(* IEC 61131-3 sources: daoli-st-library/DL_Base (part 11) *)

(* ---- FB_DL_DutyStandbyRotation.st ---- *)
(*==============================================================================
 * 组件名称 (Component)  : FB_DL_DutyStandbyRotation
 * 所属子库 (Sublibrary) : DL_Base
 * 当前版本 (Version)    : 1.0.0
 * 兼容性   (Platform)   : CODESYS 3.5 / TwinCAT 3 / 汇川 InoProShop / Machine Expert
 *                         仅依赖 Standard.library（TON / R_TRIG / ABS），零厂商方言
 * 功能描述 (Function)   : 8 台泵 / 风机 / 压缩机的主备轮值与均衡调度。
 *                         按累计运行时间排序，把"需求台数"分给运行时间最短且满足启动条件
 *                         的机组；按周期把领机降为备机、备机升为领机；故障机立即跳过；
 *                         每台机受最小运行时长与最小停机时长双重保护，避免刚启就停把
 *                         接触器打烂；任何时刻不得把在运行的机组全部停掉。
 *                         解决多泵系统两类对立顽疾："永远只跑 1 号泵、2 号泵锈死"与
 *                         "轮值切得太勤、接触器与软启动器半年一换"。
 *
 * 【安全语义 / Safety semantics（编码侧不可弱化的四条）】
 *   1) 命令-反馈分离：本块只发启动命令（cmd 语义，FALSE = 停），运行状态一律以
 *      abUnitRunning 反馈为准，绝不假设"发了命令就等于在转"。
 *   2) 先启后停：停机放行条件是"目标集中已在运行的台数 >= 需求台数"，比"在运行台数
 *      >= 需求台数"更严。后者在换机场景下仍会短暂欠载（压力/流量掉一拍），本块刻意收紧。
 *   3) 故障机越权停机：abUnitFault = TRUE 且仍在运行时立即撤销命令，越过最小运行时长。
 *      这是最小运行时长保护的唯一例外。
 *   4) 无可用机组时（需求 > 0 且可用 = 0）已在运行的机组绝不因此被停——现场可能是
 *      就地/检修状态把"就绪"信号摘掉了，停掉正在供压的泵比少启一台危险得多。
 *
 * 【失真与语义披露 / Distortion disclosure】
 *   1) 运行时间账（afRunSec / auStartCount）是否断电保持由调用方决定（Retain 声明在
 *      调用侧）。不保持则每次上电从 0 起轮，轮值顺序每次开机都从 0 号机开始。
 *   2) 时间换算按 TIME 基准 1 ms（CODESYS / TwinCAT 3 / 汇川三平台一致）。移植到
 *      100 ns 基准平台时只需改 DL_DS_MS_PER_S 处的一行换算，逻辑不动。
 *   3) 按接口契约，参数冲突故障的复位沿会清零运行时间账——等同重置最小时长约束，
 *      复位前必须确认机组处于稳定工况（手册列为操作注意事项）。
 *   4) 排序为选择排序 O(64)。同运行时间的 tie-break 取"上一拍序列位置"而非索引升序：
 *      若死守索引升序，段 7 刚做完的轮值会在下一拍重新排序时被原样排回去，轮值等于
 *      永不生效（本批实测踩到的实现陷阱）。首扫序列为 0..7 恒等排列，因此冷启动行为
 *      与"索引升序"完全一致；轮值之后同值机组按轮值后的相对顺序排列，结果仍可复算。
 *
 * 开源溯源 (Origin)     : 原创实现（参考西门子 LBP 基础过程库中"最多 8 台聚合体"的粒度
 *                         与 cmd/ind 命令-反馈分离思想，以及 lead-lag 主备轮值工艺惯例，
 *                         clean-room 编写，未接触也未复制任何 LBP 源码）
 * 本文件内含       : TYPE  E_DL_RotationState（配套枚举，归属 DL_Base）
 *                    FB    FB_DL_DutyStandbyRotation
 * 依赖     (Depends)    : 无 DL_ 内部依赖；Standard.library: TON / R_TRIG
 * 红线自检 (Redline)    : R1 ✓ 零全局变量表与外部变量引用 ｜ R2 ✓ 零物理 IO 地址直写
 *                         R3 ✓ 纯 IEC 61131-3（定长数组 + 选择排序，无动态内存）
 *                         R4 ✓ 需求钳位 + 时间增量钳位 + 双向最小时长 + 计数饱和
 *                         R5 ✓ 全变量中英双语同行注释 ｜ R6 ✓ 四态 ENUM + CASE + ELSE 兜底
 *                         R7 ✓ 三实例主体最前部无条件刷新（本组件核心考点）
 * 修订历史 (Revision)   :
 *   2026-11-14  v1.0.0  首版入库（Phase 1 收口批次 · R3）
 *============================================================================*)

(*-----------------------------------------------------------------------------
 * 枚举: E_DL_RotationState（归属 DL_Base，与 FB_DL_DutyStandbyRotation 同文件）
 * 含义: 轮值调度主状态。数值步长留空位便于后续插态而不破坏已有工程。
 *----------------------------------------------------------------------------*)
TYPE E_DL_RotationState :
(
    eIdle          := 0,     // 未使能：命令全部撤销，运行时间账继续按反馈累加 / Disabled, commands dropped, runtime still accounted
    eRunning       := 10,    // 正常调度：累加 → 排序 → 定需求集 → 先启后停 / Normal scheduling
    eRotatePending := 20,    // 轮值挂起：受最小时长阻挡，保持当前组合并每拍重试 / Rotation pending, retried every scan
    eFault         := 99     // 参数冲突锁存：轮值禁用，但启停调度照常工作 / Latched config fault, scheduling still runs
);
END_TYPE

(*==============================================================================
 * 功能块: FB_DL_DutyStandbyRotation
 * 调用约定: 每个扫描周期无条件调用一次，uDeltaTimeMs 必须注入真实任务间隔。
 *============================================================================*)
FUNCTION_BLOCK FB_DL_DutyStandbyRotation
VAR_INPUT
    abUnitReady     : ARRAY[0..7] OF BOOL;    // 机组就绪（无故障、无就地、无禁止），上限 8 台 / Unit ready, max 8 units
    abUnitRunning   : ARRAY[0..7] OF BOOL;    // 运行反馈（接触器辅助触点或流量开关）/ Running feedback
    abUnitFault     : ARRAY[0..7] OF BOOL;    // 机组故障（跳过并允许立即停机）/ Unit fault, skipped and stopped at once
    nDemand         : INT := 0;               // 需求运行台数，合法域 0..8 / Required unit count, valid 0..8
    bEnable         : BOOL := TRUE;           // 使能，FALSE 时命令全撤 / Enable, FALSE drops all commands
    uDeltaTimeMs    : UDINT;                  // 调用方注入的扫描间隔 [ms] / Injected scan delta [ms]
    tMinRunTime     : TIME := T#10M;          // 最小连续运行时长 [min]，防刚启就停 / Minimum run time
    tMinStopTime    : TIME := T#5M;           // 最小停机时长 [min]，防接触器高频动作 / Minimum stop time
    tRotateInterval : TIME := T#24H;          // 轮值周期 [h] / Rotation interval
    bForceRotate    : BOOL;                   // 上升沿：立即请求一次轮值（仍受最小时长约束）/ Rising edge: force one rotation
    bReset          : BOOL;                   // 上升沿：复位参数冲突并清零运行时间账 / Rising edge: reset the config fault and clear runtimes
END_VAR
VAR_OUTPUT
    abStartCmd        : ARRAY[0..7] OF BOOL;  // 启动命令（cmd 语义，FALSE = 停）/ Start command per unit, FALSE = stop
    anRank            : ARRAY[0..7] OF INT;   // 本轮优先顺序，0 = 最高 / Priority rank, 0 = highest
    nLeadUnit         : INT;                  // 领机号 0..7，-1 = 无 / Lead unit 0..7, -1 = none
    afRuntimeHours    : ARRAY[0..7] OF LREAL; // 累计运行小时 [h] / Accumulated runtime [h]
    abBlockedByMinRun : ARRAY[0..7] OF BOOL;  // 因最小运行时长被阻止停机 / Stop blocked by the minimum run time
    abBlockedByMinStop: ARRAY[0..7] OF BOOL;  // 因最小停机时长被阻止启动 / Start blocked by the minimum stop time
    auStartCount      : ARRAY[0..7] OF UDINT; // 各机启动次数（饱和）/ Start count per unit, saturating
    bRotatePending    : BOOL;                 // 轮值挂起中 / Rotation pending
    bNoAvailableUnit  : BOOL;                 // 无可用机组（瞬时诊断）/ No available unit, instantaneous
    uRotateCount      : UDINT;                // 已完成的轮值次数（饱和）/ Completed rotations, saturating
    bError            : BOOL;                 // 故障标志（参数冲突锁存）/ Fault flag, config conflict latched
    uErrorId          : UDINT;                // 故障码，0 = 无故障 / Error code, 0 = no error
    eState            : E_DL_RotationState;   // 当前状态（供 HMI 诊断）/ Current state for HMI diagnosis
END_VAR
VAR
    fbTrigReset     : R_TRIG;                 // 复位上升沿检测实例 / Reset rising edge detector
    fbTrigForce     : R_TRIG;                 // 强制轮值上升沿检测实例 / Force-rotate rising edge detector
    fbTonRotate     : TON;                    // 轮值周期定时器 / Rotation interval timer
    eStateInt       : E_DL_RotationState;     // 主状态机内部当前态 / Internal state of the main state machine
    afRunSec        : ARRAY[0..7] OF LREAL;   // 运行秒累加 [s] / Runtime seconds accumulator [s]
    afStopSec       : ARRAY[0..7] OF LREAL;   // 停机秒累加 [s] / Stop seconds accumulator [s]
    anOrder         : ARRAY[0..7] OF INT;     // 已提交的优先序列（可用优先，运行时间升序）/ Committed priority order
    anTrial         : ARRAY[0..7] OF INT;     // 轮值试验序列（未提交前不生效）/ Trial order, not committed yet
    anPos           : ARRAY[0..7] OF INT;     // 各机组在上一拍序列中的位置（排序稳定性锚点）/ Previous position per unit
    abUsable        : ARRAY[0..7] OF BOOL;    // 可用 = 就绪且无故障 / Usable = ready and not faulted
    abDesired       : ARRAY[0..7] OF BOOL;    // 目标运行集 / Desired running set
    abTrialUnit     : ARRAY[0..7] OF BOOL;    // 轮值试验目标集 / Trial desired set
    abCmdInt        : ARRAY[0..7] OF BOOL;    // 本拍命令内部副本 / Internal command copy of this scan
    abCmdPrev       : ARRAY[0..7] OF BOOL;    // 上一拍命令（算启动沿）/ Previous commands, for start edges
    nIdx            : INT;                    // 外层索引 / Outer index
    nInner          : INT;                    // 内层索引 / Inner index
    nMinPos         : INT;                    // 选择排序中的最小元位置 / Position of the minimum during selection sort
    nTmp            : INT;                    // 交换临时量 / Swap temporary
    nAvail          : INT;                    // 可用机组数 / Number of usable units
    nDesired        : INT;                    // 本拍应运行台数（已按可用数钳位）/ Desired count, clamped to the usable count
    nRunningCnt     : INT;                    // 当前在运行台数 / Currently running units
    nDesiredRunning : INT;                    // 目标集中已在运行的台数 / Desired units already running
    nCnt            : INT;                    // 计数累加器 / Counting accumulator
    nLead           : INT;                    // 领机号 / Lead unit index
    nDemandEff      : INT;                    // 钳位后的需求台数 / Clamped demand
    fDtSec          : LREAL;                  // 扫描间隔换算成秒 [s] / Scan delta in seconds [s]
    fMinRunSec      : LREAL;                  // 最小运行时长 [s] / Minimum run time [s]
    fMinStopSec     : LREAL;                  // 最小停机时长 [s] / Minimum stop time [s]
    tRotEff         : TIME;                   // 钳位后的轮值周期 [ms] / Clamped rotation interval [ms]
    uDtEff          : UDINT;                  // 钳位后的扫描间隔 [ms] / Clamped scan delta [ms]
    uWarnId         : UDINT;                  // 本拍瞬时告警码 / Instantaneous warning code of this scan
    uRotateCnt      : UDINT;                  // 轮值次数内部副本（饱和）/ Internal rotation counter, saturating
    bRotateReq      : BOOL;                   // 本拍请求轮值 / Rotation requested this scan
    bRotTimerRun    : BOOL;                   // 轮值定时器运行中 / Rotation timer running
    bRotTimerRearm  : BOOL;                   // 轮值定时器下一拍重新计时 / Rearm the rotation timer next scan
    bRotPendingScr  : BOOL;                   // 本拍轮值因最小时长受阻 / Rotation blocked by the minimum times this scan
    bFeasible       : BOOL;                   // 轮值试验是否可行 / Whether the trial rotation is feasible
    bSmaller        : BOOL;                   // 排序比较：候选元是否更靠前 / Sort comparator: candidate ranks earlier
    bHoldAll        : BOOL;                   // 无可用机组时冻结全部停机 / Freeze every stop when no unit is usable
    bSchedOn        : BOOL;                   // 本拍允许调度 / Scheduling enabled this scan
    bConflict       : BOOL;                   // 本拍存在时间参数冲突 / Time-parameter conflict present this scan
    bParamLatch     : BOOL;                   // 参数冲突锁存 / Configuration conflict latched
    bStateFault     : BOOL;                   // 非法状态锁存（与参数冲突分开记账）/ Illegal-state latch, kept apart from the config latch
    bCntWarned      : BOOL;                   // 饱和告警已发过一次 / Saturation warning already raised
    bSortInit       : BOOL := TRUE;           // 排序序列尚未初始化为恒等排列 / Priority order not yet initialised
    bFirstScan      : BOOL := TRUE;           // 上电首扫标志 / First-scan flag
END_VAR
VAR CONSTANT
    DL_DS_UNITS      : INT   := 8;            // 机组数，必须等于数组维度 / Unit count, must match the arrays
    DL_DS_IDX_NONE   : INT   := -1;           // 无效索引哨兵 / Invalid-index sentinel
    DL_DS_HOUR_MAX   : LREAL := 1.0E9;        // 运行小时饱和上限 [h] / Runtime saturation [h]
    DL_DS_SEC_MAX    : LREAL := 3.6E12;       // 运行秒饱和上限 [s]，与小时上限对齐 / Runtime saturation [s]
    DL_DS_SEC_PER_H  : LREAL := 3600.0;       // 小时换算常数 [s/h] / Seconds per hour
    DL_DS_MS_PER_S   : LREAL := 1000.0;       // 毫秒换算常数 [ms/s]，三平台 TIME 基准均为 1 ms / Milliseconds per second
    DL_DS_DT_MAX     : UDINT := 60000;        // 时间增量上限 [ms]，超此值判为断点 / Delta clamp [ms]
    DL_DS_EPS        : LREAL := 1.0E-6;       // 浮点判等容差 / Float comparison tolerance
    DL_DS_CNT_MAX    : UDINT := 16#FFFF_FFFE; // 计数器饱和值 / Counter saturation
    DL_DS_ROT_MIN    : TIME  := T#1S;         // 轮值周期下限 [s] / Rotation interval lower bound
    DL_DS_ROT_MAX    : TIME  := T#8760H;      // 轮值周期上限 [h]，一年 / Rotation interval upper bound
END_VAR

(*------------------------------------------------------------------------------
 * 段 0｜轮值周期钳位（先于定时器，避免 PT = 0 造成每拍触发）
 *      Rotation-interval clamp, done before the timer so PT is never zero
 *-----------------------------------------------------------------------------*)
uWarnId := 16#0000;
tRotEff := tRotateInterval;

IF tRotEff < DL_DS_ROT_MIN THEN
    tRotEff := DL_DS_ROT_MIN;
    uWarnId := 16#0001_0001;
ELSIF tRotEff > DL_DS_ROT_MAX THEN
    tRotEff := DL_DS_ROT_MAX;
    uWarnId := 16#0001_0001;
END_IF

(*------------------------------------------------------------------------------
 * 段 1｜无条件刷新区（红线 R7）：两沿 + 一轮值周期计时
 *      Unconditional refresh zone: two edges plus the rotation interval timer
 *      IN 由 bRotTimerRun 这一派生量给出，实例调用本身绝不进 IF
 *-----------------------------------------------------------------------------*)
fbTrigReset(CLK := bReset);
fbTrigForce(CLK := bForceRotate);
fbTonRotate(IN := bRotTimerRun, PT := tRotEff);

bRotateReq := fbTrigForce.Q;

IF fbTonRotate.Q THEN
    bRotateReq     := TRUE;
    bRotTimerRun   := FALSE;    // 下一拍 ET 归零 / Reset ET on the next scan
    bRotTimerRearm := TRUE;
ELSIF bRotTimerRearm THEN
    bRotTimerRun   := TRUE;
    bRotTimerRearm := FALSE;
END_IF

(*------------------------------------------------------------------------------
 * 段 2｜上电首扫：状态、领机号与锁存显式落到安全侧
 *      First-scan init: state, lead index and latches forced to the safe side
 *-----------------------------------------------------------------------------*)
IF bFirstScan THEN
    bFirstScan  := FALSE;
    eStateInt   := E_DL_RotationState.eIdle;
    nLead       := DL_DS_IDX_NONE;
    bParamLatch := FALSE;
    uRotateCnt  := 0;
    bRotTimerRun   := FALSE;
    bRotTimerRearm := TRUE;
END_IF

(*------------------------------------------------------------------------------
 * 段 3｜时间增量校验（边界 B8）：0 或超上限一律钳位，绝不接受回绕值
 *      Delta-time check: zero or over-limit values are clamped, wraparound never accepted
 *      回绕的 UDINT 转成秒后是天文数字，会瞬间把运行时间算爆并把排序彻底打乱
 *-----------------------------------------------------------------------------*)
IF uDeltaTimeMs = 0 THEN
    uDtEff  := 1;
    uWarnId := 16#0001_0008;
ELSIF uDeltaTimeMs > DL_DS_DT_MAX THEN
    uDtEff  := DL_DS_DT_MAX;
    uWarnId := 16#0001_0008;
ELSE
    uDtEff := uDeltaTimeMs;
END_IF

fDtSec     := UDINT_TO_LREAL(uDtEff) / DL_DS_MS_PER_S;
fMinRunSec := TIME_TO_LREAL(tMinRunTime) / DL_DS_MS_PER_S;
fMinStopSec := TIME_TO_LREAL(tMinStopTime) / DL_DS_MS_PER_S;

(*------------------------------------------------------------------------------
 * 段 4｜参数校验（边界 B1/B7）
 *      Parameter validation: demand clamp and the minimum-time conflict check
 *-----------------------------------------------------------------------------*)
nDemandEff := nDemand;
IF nDemand < 0 THEN
    nDemandEff := 0;
    uWarnId    := 16#0001_0001;
ELSIF nDemand > DL_DS_UNITS THEN
    nDemandEff := DL_DS_UNITS;
    uWarnId    := 16#0001_0001;
END_IF

(* 最小运行 + 最小停机 > 轮值周期：轮值永远等不到，属参数冲突而非运行故障 *)
(* min-run + min-stop > interval means rotation could never complete: a configuration conflict *)
bConflict := ((tMinRunTime + tMinStopTime) > tRotateInterval);

IF bConflict THEN
    bParamLatch := TRUE;
END_IF

IF (tMinRunTime < T#0S) OR (tMinStopTime < T#0S) THEN
    uWarnId := 16#0001_0001;
END_IF

(*------------------------------------------------------------------------------
 * 段 5｜运行时间记账（状态 eIdle 也照记：停机也要记账，否则轮值失真）
 *      Runtime accounting runs even when disabled: an unaccounted stop skews rotation
 *      以反馈为准而不是以命令为准，接触器没吸合就不能算运行
 *-----------------------------------------------------------------------------*)
FOR nIdx := 0 TO (DL_DS_UNITS - 1) DO

    IF abUnitRunning[nIdx] THEN
        afRunSec[nIdx] := afRunSec[nIdx] + fDtSec;
        IF afRunSec[nIdx] > DL_DS_SEC_MAX THEN
            afRunSec[nIdx] := DL_DS_SEC_MAX;
            uWarnId := 16#0001_0007;
        END_IF
    ELSE
        afStopSec[nIdx] := afStopSec[nIdx] + fDtSec;
        IF afStopSec[nIdx] > DL_DS_SEC_MAX THEN
            afStopSec[nIdx] := DL_DS_SEC_MAX;
        END_IF
    END_IF

    afRuntimeHours[nIdx] := afRunSec[nIdx] / DL_DS_SEC_PER_H;
    IF afRuntimeHours[nIdx] > DL_DS_HOUR_MAX THEN
        afRuntimeHours[nIdx] := DL_DS_HOUR_MAX;
    END_IF

END_FOR

(*------------------------------------------------------------------------------
 * 段 6｜可用性与候选排序（边界 B6/B10）
 *      Usability and candidate ordering: usable first, then runtime, then previous position
 *      序列只在首扫初始化为恒等排列，之后一律在既有排列上就地排序：
 *      若每拍都从 0..7 重新开始排，段 7 刚做完的轮值会在下一拍被排序抹掉，
 *      轮值等于永远不生效——这是本组件最容易踩的实现陷阱
 *      The order is initialised once and then sorted in place, otherwise every rotation
 *      would be erased by the next scan's re-sort
 *-----------------------------------------------------------------------------*)
nAvail := 0;

FOR nIdx := 0 TO (DL_DS_UNITS - 1) DO
    abUsable[nIdx] := abUnitReady[nIdx] AND (NOT abUnitFault[nIdx]);
    IF abUsable[nIdx] THEN
        nAvail := nAvail + 1;
    END_IF
END_FOR

IF bSortInit THEN
    FOR nIdx := 0 TO (DL_DS_UNITS - 1) DO
        anOrder[nIdx] := nIdx;
        anPos[nIdx]   := nIdx;
    END_FOR
    bSortInit := FALSE;
END_IF

(* 选择排序：8 元定长，0..6 外层、nIdx+1..7 内层，迭代次数由常量卡死 *)
(* Selection sort over 8 fixed elements, the loop bounds are compile-time constants *)
FOR nIdx := 0 TO (DL_DS_UNITS - 2) DO

    nMinPos := nIdx;

    FOR nInner := (nIdx + 1) TO (DL_DS_UNITS - 1) DO

        bSmaller := FALSE;

        IF abUsable[anOrder[nInner]] AND (NOT abUsable[anOrder[nMinPos]]) THEN
            bSmaller := TRUE;
        ELSIF abUsable[anOrder[nInner]] = abUsable[anOrder[nMinPos]] THEN
            IF (afRunSec[anOrder[nInner]] + DL_DS_EPS) < afRunSec[anOrder[nMinPos]] THEN
                bSmaller := TRUE;
            ELSIF ABS(afRunSec[anOrder[nInner]] - afRunSec[anOrder[nMinPos]]) <= DL_DS_EPS THEN
                (* 运行时间相同：按上一拍位置排序，保证稳定且轮值结果不被抹掉 *)
                (* Equal runtime: keep the previous relative order, so rotations survive *)
                IF anPos[anOrder[nInner]] < anPos[anOrder[nMinPos]] THEN
                    bSmaller := TRUE;
                END_IF
            END_IF
        END_IF

        IF bSmaller THEN
            nMinPos := nInner;
        END_IF

    END_FOR

    IF nMinPos <> nIdx THEN
        nTmp             := anOrder[nIdx];
        anOrder[nIdx]    := anOrder[nMinPos];
        anOrder[nMinPos] := nTmp;
    END_IF

END_FOR

FOR nIdx := 0 TO (DL_DS_UNITS - 1) DO
    anPos[anOrder[nIdx]] := nIdx;
END_FOR

nDesired := nDemandEff;
IF nDesired > nAvail THEN
    nDesired := nAvail;
END_IF

(*------------------------------------------------------------------------------
 * 段 7｜轮值尝试（边界 B7）：可行才移位，不可行一律不动任何命令
 *      Rotation attempt: shift only when every constraint is met, never touch commands otherwise
 *      把"领机移到可用序列末位、其余前移一位"这一动作做成试验序列，
 *      可行性由"要停的机组已满足最小运行、要启的机组已满足最小停机"共同决定
 *-----------------------------------------------------------------------------*)
bRotPendingScr := FALSE;

FOR nIdx := 0 TO (DL_DS_UNITS - 1) DO
    abBlockedByMinRun[nIdx]  := FALSE;
    abBlockedByMinStop[nIdx] := FALSE;
END_FOR

IF bRotateReq AND bEnable AND (NOT bParamLatch)
   AND (eStateInt <> E_DL_RotationState.eIdle)
   AND (eStateInt <> E_DL_RotationState.eFault)
   AND (nAvail >= 2) AND (nDesired >= 1) THEN

    FOR nIdx := 0 TO (DL_DS_UNITS - 1) DO
        anTrial[nIdx] := anOrder[nIdx];
    END_FOR

    nTmp := anTrial[0];
    FOR nIdx := 0 TO (DL_DS_UNITS - 2) DO
        IF nIdx < (nAvail - 1) THEN
            anTrial[nIdx] := anTrial[nIdx + 1];
        END_IF
    END_FOR
    anTrial[nAvail - 1] := nTmp;

    (* 试验目标集：可用序列中取前 nDesired 台 *)
    (* Trial set: the first nDesired usable entries of the trial order *)
    FOR nIdx := 0 TO (DL_DS_UNITS - 1) DO
        abTrialUnit[nIdx] := FALSE;
    END_FOR

    nCnt := 0;
    FOR nIdx := 0 TO (DL_DS_UNITS - 1) DO
        IF (nCnt < nDesired) AND abUsable[anTrial[nIdx]] AND (NOT abTrialUnit[anTrial[nIdx]]) THEN
            abTrialUnit[anTrial[nIdx]] := TRUE;
            nCnt := nCnt + 1;
        END_IF
    END_FOR

    (* 可行性检查：需停的看最小运行，需启的看最小停机；故障机不参与（越权立即停） *)
    (* Feasibility: stops need the min run time, starts need the min stop time *)
    bFeasible := TRUE;

    FOR nIdx := 0 TO (DL_DS_UNITS - 1) DO
        IF abUnitRunning[nIdx] AND (NOT abTrialUnit[nIdx]) AND (NOT abUnitFault[nIdx]) THEN
            IF afRunSec[nIdx] < fMinRunSec THEN
                bFeasible := FALSE;
                abBlockedByMinRun[nIdx] := TRUE;
            END_IF
        END_IF
        IF (NOT abUnitRunning[nIdx]) AND abTrialUnit[nIdx] THEN
            IF afStopSec[nIdx] < fMinStopSec THEN
                bFeasible := FALSE;
                abBlockedByMinStop[nIdx] := TRUE;
            END_IF
        END_IF
    END_FOR

    IF bFeasible THEN
        FOR nIdx := 0 TO (DL_DS_UNITS - 1) DO
            anOrder[nIdx] := anTrial[nIdx];
        END_FOR
        (* 提交后立即刷新位置锚点，否则下一次排序会按旧位置把轮值结果排回去 *)
        (* Refresh the position anchor at once, or the next sort undoes the rotation *)
        FOR nIdx := 0 TO (DL_DS_UNITS - 1) DO
            anPos[anOrder[nIdx]] := nIdx;
        END_FOR
        bRotateReq := FALSE;
        IF uRotateCnt < DL_DS_CNT_MAX THEN
            uRotateCnt := uRotateCnt + 1;
        ELSIF NOT bCntWarned THEN
            uWarnId    := 16#0001_0007;
            bCntWarned := TRUE;
        END_IF
    ELSE
        (* 边界 B7：请求不丢，保留到条件满足，每拍重试且只补做一次 *)
        (* The request is kept, retried every scan, and only ever executed once *)
        bRotPendingScr := TRUE;
    END_IF

END_IF

(*------------------------------------------------------------------------------
 * 段 8｜主状态机（红线 R6）：ENUM + CASE + ELSE 兜底
 *      Main state machine with the mandatory ELSE fallback
 *-----------------------------------------------------------------------------*)
CASE eStateInt OF

    E_DL_RotationState.eIdle:
        bRotateReq     := FALSE;
        bRotTimerRun   := FALSE;
        bRotTimerRearm := TRUE;
        IF bEnable THEN
            IF bParamLatch THEN
                eStateInt := E_DL_RotationState.eFault;
            ELSE
                eStateInt := E_DL_RotationState.eRunning;
            END_IF
        END_IF

    E_DL_RotationState.eRunning:
        IF NOT bEnable THEN
            eStateInt := E_DL_RotationState.eIdle;
        ELSIF bParamLatch THEN
            eStateInt := E_DL_RotationState.eFault;
        ELSIF bRotPendingScr THEN
            eStateInt := E_DL_RotationState.eRotatePending;
        END_IF

    E_DL_RotationState.eRotatePending:
        IF NOT bEnable THEN
            eStateInt := E_DL_RotationState.eIdle;
        ELSIF bParamLatch THEN
            eStateInt := E_DL_RotationState.eFault;
        ELSIF NOT bRotPendingScr THEN
            eStateInt := E_DL_RotationState.eRunning;
        END_IF

    E_DL_RotationState.eFault:
        (* 轮值禁用但启停调度照常：不能因为轮值配错就让泵不转 *)
        (* Rotation is disabled, scheduling still runs: a wrong interval must not stop the pumps *)
        bRotateReq := FALSE;
        IF NOT bEnable THEN
            eStateInt := E_DL_RotationState.eIdle;
        ELSIF fbTrigReset.Q AND (NOT bConflict) THEN
            bParamLatch := FALSE;
            bStateFault := FALSE;
            eStateInt   := E_DL_RotationState.eRunning;
            (* 接口契约：复位参数冲突同时清零运行时间账，等同重置最小时长约束 *)
            (* Contract: resetting the conflict also clears the runtime books *)
            FOR nIdx := 0 TO (DL_DS_UNITS - 1) DO
                afRunSec[nIdx]    := 0.0;
                afStopSec[nIdx]   := 0.0;
                afRuntimeHours[nIdx] := 0.0;
            END_FOR
            bRotTimerRun   := FALSE;
            bRotTimerRearm := TRUE;
        END_IF

    ELSE
        (* 非法状态拦截：不做隐式恢复，直接锁存上报 *)
        (* Illegal state interception: no implicit recovery, latch and report *)
        eStateInt   := E_DL_RotationState.eFault;
        bStateFault := TRUE;

END_CASE;

bSchedOn := bEnable AND (eStateInt <> E_DL_RotationState.eIdle);

(*------------------------------------------------------------------------------
 * 段 9｜命令生成（边界 B1/B2/B3/B4/B5）：先启后停，单一出口
 *      Command derivation: starts first, stops last, single exit
 *      顺序本身即安全逻辑：先把替代机组拉起来，等反馈确认到位后才允许停旧机
 *-----------------------------------------------------------------------------*)
FOR nIdx := 0 TO (DL_DS_UNITS - 1) DO
    abDesired[nIdx] := FALSE;
END_FOR

nCnt := 0;
FOR nIdx := 0 TO (DL_DS_UNITS - 1) DO
    IF (nCnt < nDesired) AND abUsable[anOrder[nIdx]] THEN
        abDesired[anOrder[nIdx]] := TRUE;
        nCnt := nCnt + 1;
    END_IF
END_FOR

nRunningCnt     := 0;
nDesiredRunning := 0;

FOR nIdx := 0 TO (DL_DS_UNITS - 1) DO
    IF abUnitRunning[nIdx] THEN
        nRunningCnt := nRunningCnt + 1;
        IF abDesired[nIdx] THEN
            nDesiredRunning := nDesiredRunning + 1;
        END_IF
    END_IF
END_FOR

(* 边界 B1/V5：需求 > 0 而可用 = 0 时冻结全部停机，已在供压的机组绝不停 *)
(* Demand > 0 with no usable unit freezes every stop: a running pump is never stopped *)
bHoldAll := (nDemandEff > 0) AND (nAvail = 0);

FOR nIdx := 0 TO (DL_DS_UNITS - 1) DO

    abCmdInt[nIdx] := abDesired[nIdx];

    IF abUnitFault[nIdx] THEN
        (* 边界 B4：故障机越权停机，不等最小运行时长 *)
        (* Fault overrides the minimum run time: stop at once *)
        abCmdInt[nIdx] := FALSE;

    ELSIF abDesired[nIdx] AND (NOT abUnitRunning[nIdx]) THEN
        (* 启动约束：未就绪或停机未满，一律不启动 *)
        (* Start constraint: not ready or the minimum stop time is not satisfied *)
        IF (NOT abUnitReady[nIdx]) THEN
            abCmdInt[nIdx] := FALSE;
        ELSIF afStopSec[nIdx] < fMinStopSec THEN
            abCmdInt[nIdx] := FALSE;
            abBlockedByMinStop[nIdx] := TRUE;
        END_IF

    ELSIF abUnitRunning[nIdx] AND (NOT abDesired[nIdx]) THEN
        (* 停机约束：冻结 → 最后一台 → 最小运行时长 → 目标集是否已全部到位 *)
        (* Stop constraint: freeze, then the last unit, then min run, then start-first *)
        IF bHoldAll THEN
            abCmdInt[nIdx] := TRUE;
        ELSIF (nDemandEff > 0) AND (nRunningCnt <= 1) THEN
            (* 边界 B5 加强项：需求 > 0 时绝不停掉正在供压的最后一台 *)
            (* Never stop the last running unit while a demand exists *)
            abCmdInt[nIdx] := TRUE;
        ELSIF afRunSec[nIdx] < fMinRunSec THEN
            abCmdInt[nIdx] := TRUE;
            abBlockedByMinRun[nIdx] := TRUE;
        ELSIF nDesiredRunning >= nDesired THEN
            abCmdInt[nIdx] := FALSE;
        ELSE
            abCmdInt[nIdx] := TRUE;
        END_IF

    END_IF

END_FOR

IF NOT bSchedOn THEN
    FOR nIdx := 0 TO (DL_DS_UNITS - 1) DO
        abCmdInt[nIdx] := FALSE;
    END_FOR
END_IF

(*------------------------------------------------------------------------------
 * 段 10｜启动次数统计（命令上升沿）：饱和累加，回绕会让保养周期判断失效
 *      Start counters increment on command rising edges, with saturation
 *-----------------------------------------------------------------------------*)
FOR nIdx := 0 TO (DL_DS_UNITS - 1) DO
    IF abCmdInt[nIdx] AND (NOT abCmdPrev[nIdx]) THEN
        IF auStartCount[nIdx] < DL_DS_CNT_MAX THEN
            auStartCount[nIdx] := auStartCount[nIdx] + 1;
        ELSIF NOT bCntWarned THEN
            uWarnId    := 16#0001_0007;
            bCntWarned := TRUE;
        END_IF
    END_IF
    abCmdPrev[nIdx] := abCmdInt[nIdx];
END_FOR

(*------------------------------------------------------------------------------
 * 段 11｜排序与领机（边界 B6）：排名来自已提交序列，不来自本拍临时计算
 *      Ranking and lead unit come from the committed order
 *-----------------------------------------------------------------------------*)
FOR nIdx := 0 TO (DL_DS_UNITS - 1) DO
    anRank[nIdx] := DL_DS_IDX_NONE;
END_FOR

FOR nIdx := 0 TO (DL_DS_UNITS - 1) DO
    IF (anOrder[nIdx] >= 0) AND (anOrder[nIdx] < DL_DS_UNITS) THEN
        anRank[anOrder[nIdx]] := nIdx;
    END_IF
END_FOR

IF (nAvail > 0) AND (nDesired > 0) THEN
    nLead := anOrder[0];
ELSE
    nLead := DL_DS_IDX_NONE;
END_IF

(*------------------------------------------------------------------------------
 * 段 12｜故障码落码（红线 R15）：锁存码优先，瞬时码条件消失即归零
 *      Error-code policy: latched codes win, instantaneous codes clear themselves
 *-----------------------------------------------------------------------------*)
IF (nDemandEff > 0) AND (nAvail = 0) THEN
    uWarnId := 16#0002_0007;
END_IF

IF eStateInt <> E_DL_RotationState.eFault THEN
    IF uWarnId <> 16#0000 THEN
        uErrorId := uWarnId;
    ELSE
        uErrorId := 16#0000_0000;
    END_IF
END_IF

IF bParamLatch THEN
    uErrorId := 16#0002_0008;
ELSIF bStateFault THEN
    uErrorId := 16#0001_0005;
END_IF

(*------------------------------------------------------------------------------
 * 段 13｜输出单一出口（范式 P-05）
 *      Single output exit: the command array is written exactly once, here
 *-----------------------------------------------------------------------------*)
FOR nIdx := 0 TO (DL_DS_UNITS - 1) DO
    abStartCmd[nIdx] := abCmdInt[nIdx];
END_FOR

bRotatePending   := (eStateInt = E_DL_RotationState.eRotatePending);
bNoAvailableUnit := (nDemandEff > 0) AND (nAvail = 0);
uRotateCount     := uRotateCnt;
nLeadUnit        := nLead;
bError           := bParamLatch OR bStateFault;
eState           := eStateInt;
END_FUNCTION_BLOCK

(* ---- FB_DL_EdgeDivider.st ---- *)
(*
    FB_DL_EdgeDivider —— 输入沿 1/N 分频
    ------------------------------------------------------------------
    分类      : DL_Base / Signal
    前缀      : FB_DL_
    版本      : 1.0.0
    溯源      : T0-1 双稳态 / 边沿族变体（源矩阵明列「主从沿 / 分频变体」为未挖扩产点）；
                只借「分频属边沿处理族」的分类事实，分频结构、钳位与回绕纪律
                100% 自有；clean-room 重写，未复制任何闭源厂商源码，
                参考实现仅限 MIT/Apache 许可
    平台      : 纯 IEC 61131-3，CODESYS V3.5+ / TwinCAT 3 / InoProShop 通用
    作者      : 道莅代码库 · PLC编程专家（R18）
    ------------------------------------------------------------------
    功能说明  : 输入每 N 个上升沿输出一个单周期脉冲，用于「双作用气缸交替动作」
                「分料器奇偶道切换」「主轴每 N 转喷一次油」等现场语义；
                bDutyHalf 为 TRUE 且 N 为偶数时输出方波（N/2 拍高 / N/2 拍低），
                N 为奇数时退化为单拍脉冲并置信息码，绝不报故障；
                计数回绕用「比较 + 赋值」，禁用取余（三平台对负数取余不一致）；
                uPulseCnt 饱和不回绕，长期运行不会翻转。
    错误码    : 16#0001_0239 分频比超上限已钳位，或奇数 N 请求方波已退化单拍——信息级，正常防御
                16#0001_023A 预留禁用（信息级，不得挪用）
                16#0001_030C uDivide = 0，输出强制 FALSE——故障级，不做取余
                16#0001_030D 预留禁用（故障级，不得挪用）
                16#0001_030E 预留禁用（故障级，不得挪用）
    码位总账  : 16#0001_0239 用 / 16#0001_023A 预留 ｜ 16#0001_030C 用 / 16#0001_030D 预留 / 16#0001_030E 预留
    状态机    : 无 CASE，相位由 uCntInt 一个整数承载，非法状态不可能出现
    采样约定  : fbTrigIn / fbTrigPhase 在本体首部无条件刷新；输入脉宽小于一个扫描
                周期不可见，高频输入须先由硬件计数模块预处理。
    修订记录  : 2026-11-16 v1.0.0 首次入库（R18）
*)
FUNCTION_BLOCK FB_DL_EdgeDivider
VAR_INPUT
    bEnable     : BOOL;                        // 使能，FALSE 计数冻结并清输出 / enable, FALSE freezes the count and clears the output
    bIn         : BOOL;                        // 待分频信号，上升沿有效 / signal to divide, rising edge effective
    uDivide     : UINT := 2;                   // 分频比 N [倍]，范围 1~1000，1 = 直通 / division ratio N [x], range 1~1000, 1 = pass-through
    bPhaseReset : BOOL;                        // 相位复位，上升沿把计数与输出相位归零 / phase reset, rising edge zeroes the count and the output phase
    bDutyHalf   : BOOL := FALSE;               // TRUE 且 N 为偶数时输出方波 / FALSE 输出单拍脉冲 / TRUE gives a square wave on even N, FALSE gives a one-cycle pulse
END_VAR
VAR_OUTPUT
    bOut      : BOOL;                          // 分频输出 / divided output
    uCounter  : UINT;                          // 当前计数 0~N-1 [拍] / current counter 0~N-1 [cycle]
    uPulseCnt : UDINT;                         // 累计输出脉冲数，饱和计数 [次] / accumulated output pulses, saturating [times]
    eErr      : UDINT;                         // 错误码，0=正常 / error id, 0=ok
    bError    : BOOL;                          // 故障标志，eErr 为故障级时 TRUE / error flag, TRUE on fault-level eErr
END_VAR
VAR
    fbTrigIn    : R_TRIG;                      // 输入沿检测实例，本体首部无条件刷新 / input edge instance, refreshed unconditionally
    fbTrigPhase : R_TRIG;                      // 相位复位沿检测实例，本体首部无条件刷新 / phase reset edge instance, refreshed unconditionally
    bInit       : BOOL := FALSE;               // 首扫标志，初值 FALSE，判据 NOT bInit / first-scan flag, initial FALSE, tested with NOT
    uCntInt     : UINT;                        // 内部相位计数 0~N-1 [拍] / internal phase counter 0~N-1 [cycle]
    uDivEff     : UINT;                        // 生效分频比，钳位后使用 [倍] / effective ratio after clamping [x]
    bHalfMode   : BOOL;                        // 方波模式有效标志（N 为偶数时成立）/ square wave mode valid flag, only on even N
    bPulseOne   : BOOL;                        // 单拍脉冲标志，用后即清 / one-cycle pulse flag, cleared after use
END_VAR
VAR CONSTANT
    DL_DIV_MAX     : UINT := 1000;             // 分频比上限 [倍] / division ratio upper bound [x]
    DL_DIV_CNT_MAX : UDINT := 16#FFFF_FFFE;    // 脉冲计数饱和值，防回绕 [次] / pulse counter saturation value, no wrap-around [times]
    DL_DIV_HALF    : UINT := 2;                // 偶数判定与半相位除数 [无量纲] / divisor for the even check and the half phase [dimensionless]
END_VAR

// 段 1｜输出与错误状态预置 / segment 1, preset outputs and error status
bOut := FALSE;                                 // 输出先清零 / clear the output first
eErr := 0;                                     // 预置无错误 / preset no error
bError := FALSE;                               // 预置无故障 / preset no fault

// 段 2｜边沿实例无条件周期刷新（红线：严禁放入条件分支）/ segment 2, unconditional edge refresh
fbTrigIn(CLK := bIn);                          // 输入沿 / input edge
fbTrigPhase(CLK := bPhaseReset);               // 相位复位沿 / phase reset edge

// 段 3｜首扫初始化（初值 FALSE，判据 NOT bInit）/ segment 3, first-scan initialisation
IF NOT bInit THEN
    uCntInt := 0;                              // 相位从 0 起 / phase starts at zero
    bPulseOne := FALSE;                        // 单拍标志清零 / clear the one-cycle flag
    bInit := TRUE;                             // 首扫只做一次 / first scan runs once only
END_IF

// 段 4｜使能闸：冻结计数并清输出 / segment 4, enable gate freezes the counter
IF NOT bEnable THEN
    uCntInt := 0;                              // 相位归零 / phase to zero
    bPulseOne := FALSE;                        // 清单拍标志 / clear the one-cycle flag
    uCounter := 0;                             // 对外计数清零 / clear the published counter
    RETURN;                                    // 失能即出口 / disabled is the exit
END_IF

// 段 5｜分频比闸：0 为故障（不做取余），超上限先钳位 / segment 5, division ratio gate
IF uDivide < 1 THEN
    eErr := 16#0001_030C;                      // 分频比为 0 故障码 / zero ratio fault id
    bError := TRUE;                            // 置故障标志 / raise the error flag
    uCounter := 0;                             // 计数回安全值 / counter to the safe value
    RETURN;                                    // 故障级提前返回 / early return on fault
END_IF
uDivEff := uDivide;                            // 默认沿用输入值 / default to the input value
IF uDivide > DL_DIV_MAX THEN
    uDivEff := DL_DIV_MAX;                     // 超上限钳位 / clamp to the upper bound
    eErr := 16#0001_0239;                      // 钳位提示（信息级不置故障）/ clamp hint, info level never raises a fault
END_IF

// 段 6｜方波可用性判定：偶数用「半值乘二回比」，全程不用取余 / segment 6, square wave availability without any modulo
bHalfMode := FALSE;                            // 先按单拍脉冲模式 / assume the one-cycle pulse mode
IF bDutyHalf AND (uDivEff > 1) THEN
    IF ((uDivEff / DL_DIV_HALF) * DL_DIV_HALF) = uDivEff THEN
        bHalfMode := TRUE;                     // 偶数成立，方波可用 / even ratio, square wave is available
    ELSE
        eErr := 16#0001_0239;                  // 奇数 N 请求方波，退化单拍（信息级）/ odd ratio asked for a square wave, degraded to a pulse (info level)
    END_IF
END_IF

// 段 7｜相位复位（优先于计数）/ segment 7, phase reset has priority over counting
IF fbTrigPhase.Q THEN
    uCntInt := 0;                              // 相位归零 / phase to zero
    bPulseOne := FALSE;                        // 复位拍不出脉冲，防自杀 / no pulse on the reset cycle, prevents self-kill
END_IF

// 段 8｜N = 1 直通模式 / segment 8, pass-through mode when N equals 1
IF uDivEff <= 1 THEN
    bOut := bIn;                               // 直通输出 / pass the input straight through
    uCntInt := 0;                              // 直通不累计相位 / no phase accumulation in pass-through
    uCounter := 0;                             // 对外计数归零 / publish a zero counter
    RETURN;                                    // 直通即出口 / pass-through is the exit
END_IF

// 段 9｜计数与回绕（比较 + 赋值，禁用取余）/ segment 9, counting and wrap-around by compare-and-assign
IF fbTrigIn.Q THEN
    uCntInt := uCntInt + 1;                    // 每个输入沿相位加一 / one phase step per input edge
    IF uCntInt >= uDivEff THEN
        uCntInt := 0;                          // 到达 N 即回零 / wrap to zero when reaching N
        bPulseOne := TRUE;                     // 跳变拍产生单拍脉冲 / the wrap cycle produces a one-cycle pulse
        IF uPulseCnt < DL_DIV_CNT_MAX THEN
            uPulseCnt := uPulseCnt + 1;        // 饱和加一，绝不回绕 / saturating increment, never wraps
        END_IF
    END_IF
END_IF

// 段 10｜输出形态：方波由相位直接派生，单拍脉冲用后即清（保持量另立变量）/ segment 10, output shape
IF bHalfMode THEN
    IF uCntInt >= (uDivEff / DL_DIV_HALF) THEN
        bOut := TRUE;                          // 后半相位为高 / high during the second half of the phase
    ELSE
        bOut := FALSE;                         // 前半相位为低 / low during the first half of the phase
    END_IF
ELSE
    bOut := bPulseOne;                         // 单拍模式直接镜像脉冲标志 / mirror the one-cycle flag
END_IF
bPulseOne := FALSE;                            // 用后即清，绝不跨拍残留 / consumed and cleared, never leaks to the next cycle
uCounter := uCntInt;                           // 对外镜像相位计数 / publish the phase counter
END_FUNCTION_BLOCK

(* ---- FB_DL_EdgeIntervalMeter.st ---- *)
(*
  Name        : FB_DL_EdgeIntervalMeter
  Category    : DL_Base
  Version     : 1.0.0
  Purpose     : 双沿间隔/周期/占空比测量：以自复位自由计时器逐拍累计时基，上升沿与下降沿分别测周期与高电平宽度，附抖动（间隔一阶绝对偏差 EMA）与无沿超时判据；/ Measure edge interval, period and duty cycle via a self-resetting free-running time base, with jitter (EMA of absolute interval deviation) and a no-edge timeout verdict
  溯源        : 借 t2-1-lgf·dateandtimer 的分类/参数域组织，clean-room 实现
  Boundary    : ① 时基委托：tonFree 为 1 天 PT 的自复位自由计时器（IN := NOT tonFree.Q，R188），逐拍取 ET 差分累加；跨 1 天回卷那拍差分为负 → 钳 0，单拍损失已声明；
                ② 占空比除子闸：周期 <= eps → 占空比按 0 处理（不产生 Inf）；
                ③ 无沿判据用 TIME 直比（tTimeout > 0 已过组态闸），不额外占定时器实例；
                ④ 高电平宽度为「最近一次采样值」，下降沿那拍取上拍快照（一拍滞后已在头注释声明）；
                ⑤ 计数饱和：UDINT 到上限前停加，防回绕。
*)
TYPE E_DL_EimState :
(
    eIdle  := 0,                             (* 未使能 / Disabled *)
    eRun   := 10,                            (* 测量运行 / Measuring *)
    eFault := 90                             (* 故障锁存相 / Fault latched *)
);
END_TYPE

TYPE E_DL_EimCause :
(
    eNone       := 0,                        (* 无故障成因 / No cause *)
    eCfgIllegal := 1,                        (* 组态非法：超时/扫描周期非正 / Illegal config *)
    ePhaseBad   := 2                         (* 非法相位兜底 / Illegal phase fallback *)
);
END_TYPE

FUNCTION_BLOCK FB_DL_EdgeIntervalMeter
VAR_INPUT
    bSignal   : BOOL := FALSE;               (* 被测数字信号 [-] / Monitored digital signal *)
    tTimeout  : TIME := T#5S;                (* 无沿超时判据，域 > T#0S [ms] / No-edge timeout, must be > 0 *)
    bEnable   : BOOL := TRUE;                (* 测量使能 [-] / Enable *)
    bReset    : BOOL := FALSE;               (* 复位命令，上升沿清全部统计与故障 [-] / Reset command *)
END_VAR
VAR_OUTPUT
    tInterval    : TIME;                     (* 最近一次上升沿间隔（周期）[ms] / Latest rising-to-rising interval *)
    tPulseWidth  : TIME;                     (* 最近一次高电平宽度（下降沿锁存）[ms] / Latest high pulse width, latched on falling *)
    fDuty        : REAL;                     (* 占空比 = 高宽 / 周期，域 0..1 [-] / Duty cycle, 0..1 *)
    fJitterMs    : REAL;                     (* 间隔抖动（绝对偏差 EMA）[ms] / Interval jitter, EMA of abs deviation *)
    tIntervalMin : TIME;                     (* 窗口最小间隔（本测量生命周期）[ms] / Minimum interval seen *)
    tIntervalMax : TIME;                     (* 窗口最大间隔（本测量生命周期）[ms] / Maximum interval seen *)
    bNoEdge      : BOOL;                     (* 超时无沿指示 [-] / No-edge timeout indicator *)
    nEdgeCnt     : UDINT;                    (* 累计上升沿数（饱和）[-] / Rising edge count, saturated *)
    eState       : E_DL_EimState;            (* 状态出口 / State outlet *)
    eCause       : E_DL_EimCause;            (* 故障成因出口（R190 归因唯一） / Fault cause outlet *)
    bError       : BOOL;                     (* 故障锁存标志 [-] / Fault latch flag *)
END_VAR
VAR
    _eState    : E_DL_EimState := E_DL_EimState.eIdle;   (* 内部相位（CASE 唯一写入目标） / Internal phase *)
    _eCause    : E_DL_EimCause := E_DL_EimCause.eNone;   (* 故障成因锁存量 / Latched cause *)
    rtSig      : R_TRIG;                     (* 上升沿实例，段 0 无条件调用 / Rising edge instance *)
    ftSig      : F_TRIG;                     (* 下降沿实例，段 0 无条件调用 / Falling edge instance *)
    rtReset    : R_TRIG;                     (* 复位沿实例，段 0 无条件调用 / Reset edge instance *)
    tonFree    : TON;                        (* 自由跑时基（PT = 1 天，自复位） / Free-running time base *)
    _tFreePrev : TIME;                       (* 上拍自由时基 ET 快照（差分用）[ms] / Previous free ET snapshot *)
    _tDelta    : TIME;                       (* 本拍时基增量（回卷拍钳 0）[ms] / This-scan time delta *)
    _tSinceEdge: TIME;                       (* 距上次上升沿的累计时长 [ms] / Accumulated time since last rise *)
    _tHighLive : TIME;                       (* 高电平宽度实时值（下降沿取快照）[ms] / Live high width, snapshotted on fall *)
    _tPrevInt  : TIME;                       (* 上一次间隔（抖动基准）[ms] / Previous interval for jitter *)
    _fDev      : REAL;                       (* 本次间隔绝对偏差 [ms] / Absolute interval deviation *)
    _t0        : TIME;                       (* 时间零常量（比较基准）[ms] / Time zero constant *)
    _bFault    : BOOL;                       (* 故障锁存位 / Latched fault bit *)
    _bCfgBad   : BOOL;                       (* 组态非法当拍量 / Illegal config this scan *)
    _bFinite   : BOOL;                       (* 信号有效标志（BOOL 入参恒有限，语义占位）[-] / Signal validity placeholder *)
END_VAR
VAR CONSTANT
    DL_EIM_EPS    : REAL  := 1.0E-6;         (* 除零判零容差（REAL 量级）[-] / Division epsilon *)
    DL_EIM_DAY    : TIME  := T#1D;           (* 自由时基自复位周期（1 天）[ms] / Free base period *)
    DL_EIM_CNTMAX : UDINT := 4294967295;     (* 沿计数饱和上限（R28）[-] / Edge count saturation cap *)
    DL_EIM_JITW   : REAL  := 0.3;            (* 抖动 EMA 新值权重 [-] / Jitter EMA new-sample weight *)
END_VAR

(* —— 段 0：当拍判据派生 + 实例无条件刷新（R228A；定时器/沿实例全在段 0，无 IF 包裹） —— *)
_bCfgBad := NOT (tTimeout > T#0S);                                             (* 组态闸：超时须为正（TIME 比较，无浮点） / Config gate *)
rtReset(CLK := bReset);                                                        (* 复位沿每拍必调 / Reset edge every scan *)
rtSig(CLK := bSignal);                                                         (* 上升沿每拍必调 / Rising edge every scan *)
ftSig(CLK := bSignal);                                                         (* 下降沿每拍必调 / Falling edge every scan *)
tonFree(IN := NOT tonFree.Q, PT := DL_EIM_DAY);                                (* 自由时基自复位（R188，禁外部沿清零） / Self-resetting free base *)
_tDelta := tonFree.ET - _tFreePrev;                                            (* 时基差分（ET 单调增，回卷拍为负） / Time delta *)
IF _tDelta < _t0 THEN
    _tDelta := _t0;                                                            (* 回卷拍差分为负：钳 0（单拍损失已声明） / Wrap: clamp to zero *)
END_IF
_tFreePrev := tonFree.ET;                                                      (* 本拍快照留给下拍差分 / Snapshot for next scan *)

(* —— 段 1：单拍量预清零（R107） —— *)
_bFinite := TRUE;                                                              (* BOOL 入参恒有限（语义占位，保持全路径赋值） / Always finite *)
bNoEdge := FALSE;                                                              (* 无沿指示预清，仅运行相置位 / No-edge preset *)

(* —— 段 2：复位沿处理（作用域：清故障 + 清全部统计 + 清时基 + 迁 eIdle，R283 逐项声明） —— *)
IF rtReset.Q THEN
    _bFault := FALSE;                                                          (* 清故障锁存 / Clear fault *)
    _eCause := E_DL_EimCause.eNone;                                            (* 清成因 / Clear cause *)
    tInterval := T#0S;                                                         (* 清间隔 / Clear interval *)
    tPulseWidth := T#0S;                                                       (* 清高宽 / Clear pulse width *)
    fDuty := 0.0;                                                              (* 清占空比 / Clear duty *)
    fJitterMs := 0.0;                                                          (* 清抖动 / Clear jitter *)
    tIntervalMin := T#0S;                                                      (* 清最小值 / Clear minimum *)
    tIntervalMax := T#0S;                                                      (* 清最大值 / Clear maximum *)
    nEdgeCnt := 0;                                                             (* 清沿计数 / Clear edge count *)
    _tSinceEdge := T#0S;                                                       (* 清距沿时长 / Clear since-edge *)
    _tHighLive := T#0S;                                                        (* 清高宽实时值 / Clear live width *)
    _tPrevInt := T#0S;                                                         (* 清抖动基准 / Clear jitter base *)
    _eState := E_DL_EimState.eIdle;                                            (* 迁未使能相 / Back to idle *)
END_IF

(* —— 段 3：组态故障锁存（锁存至复位沿，R189；故障相不按当下输入重推码） —— *)
IF _bCfgBad AND NOT _bFault THEN
    _bFault := TRUE;                                                           (* 锁存故障位 / Latch fault *)
    _eCause := E_DL_EimCause.eCfgIllegal;                                      (* 成因：组态非法 / Cause: illegal config *)
    _eState := E_DL_EimState.eFault;                                           (* 同步迁故障相 / Migrate to fault *)
END_IF

(* —— 段 4：CASE 主状态机（ELSE 兜底迁 eFault，红线 6） —— *)
CASE _eState OF
    E_DL_EimState.eIdle:                                                       (* 未使能：时基清零，出口保持 0 / Disabled *)
        _tSinceEdge := T#0S;                                                   (* 距沿时长清零（失能即无测量语义） / Since-edge cleared *)
        IF bEnable AND NOT _bFault THEN
            _eState := E_DL_EimState.eRun;                                     (* 使能进入测量 / Enter measuring *)
        END_IF
    E_DL_EimState.eRun:                                                        (* 测量相：时基累加 + 双沿派生 / Measuring *)
        IF NOT bEnable THEN
            _eState := E_DL_EimState.eIdle;                                    (* 失能回未使能 / Back to idle *)
        ELSE
            _tSinceEdge := _tSinceEdge + _tDelta;                              (* 距沿时长累加（本拍增量已钳非负） / Accumulate *)
            IF bSignal THEN
                _tHighLive := _tHighLive + _tDelta;                            (* 高电平期间累积宽度 / Accumulate high width *)
            END_IF
            IF rtSig.Q THEN                                                    (* 上升沿：结算一个完整周期 / Rising edge: close one period *)
                tInterval := _tSinceEdge;                                      (* 本周期 = 距上次上升沿时长 [ms] / Period *)
                IF (nEdgeCnt > 0) AND (tInterval > T#0S) THEN
                    IF (tIntervalMin = T#0S) OR (tInterval < tIntervalMin) THEN
                        tIntervalMin := tInterval;                             (* 最小值更新（首值直取） / Update minimum *)
                    END_IF
                    IF tInterval > tIntervalMax THEN
                        tIntervalMax := tInterval;                             (* 最大值更新 / Update maximum *)
                    END_IF
                    _fDev := ABS(TIME_TO_LREAL(tInterval) - TIME_TO_LREAL(_tPrevInt));   (* 绝对偏差 [ms] / Absolute deviation *)
                    fJitterMs := DL_EIM_JITW * _fDev + (1.0 - DL_EIM_JITW) * fJitterMs;  (* 抖动 EMA（系数和 = 1，无漂移） / Jitter EMA *)
                END_IF
                _tPrevInt := tInterval;                                        (* 抖动基准更新 / Jitter base update *)
                _tSinceEdge := T#0S;                                           (* 距沿时长重新起算 / Restart since-edge *)
                _tHighLive := T#0S;                                            (* 新高电平段起算 / Restart high width *)
                IF nEdgeCnt < DL_EIM_CNTMAX THEN
                    nEdgeCnt := nEdgeCnt + 1;                                  (* 沿计数饱和累加 / Saturating count *)
                END_IF
                bNoEdge := FALSE;                                              (* 有沿即清超时 / Edge clears timeout *)
            END_IF
            IF ftSig.Q THEN                                                    (* 下降沿：锁存高宽（取上拍实时快照，一拍滞后） / Falling: latch width *)
                tPulseWidth := _tHighLive;                                     (* 高电平宽度锁存 [ms] / Latch width *)
                IF tInterval > T#0S THEN
                    fDuty := TIME_TO_LREAL(tPulseWidth) / TIME_TO_LREAL(tInterval);   (* 占空比：除子已判正 [0..1] / Duty, divisor gated *)
                    IF fDuty > 1.0 THEN
                        fDuty := 1.0;                                          (* 上限饱和 1.0（量测噪声防越界） / Clamp to 1.0 *)
                    ELSIF fDuty < 0.0 THEN
                        fDuty := 0.0;                                          (* 下限饱和 0.0 / Clamp to 0.0 *)
                    END_IF
                ELSE
                    fDuty := 0.0;                                              (* 周期未建立：占空比按 0（边界②） / No period yet: duty 0 *)
                END_IF
            END_IF
            IF _tSinceEdge > tTimeout THEN
                bNoEdge := TRUE;                                               (* 超时无沿判据（TIME 直比，除子无风险） / No-edge timeout *)
            END_IF
        END_IF
    E_DL_EimState.eFault:                                                      (* 故障相：冻结保持末值，仅复位沿出 / Fault *)
        ;                                                                      (* 锁存回放（R28） / Replay from latch *)
    ELSE                                                                       (* 非法相位兜底迁安全态 / Illegal phase fallback *)
        _eState := E_DL_EimState.eFault;                                       (* 迁故障相 / To fault *)
        _bFault := TRUE;                                                       (* 同步锁存 / Latch *)
        _eCause := E_DL_EimCause.ePhaseBad;                                    (* 成因：非法相位 / Cause: illegal phase *)
END_CASE

(* —— 段 5：出口映射（bError/eState 同源，R191） —— *)
bError := _bFault;                                                             (* 故障标志镜像 / Fault flag mirror *)
eState := _eState;                                                             (* 状态出口 / State outlet *)
eCause := _eCause;                                                             (* 成因出口 / Cause outlet *)
END_FUNCTION_BLOCK

(* ---- FB_DL_EdgeMasterSlaveSync.st ---- *)
(*
  ==================================================================
  组件名 Component  : FB_DL_EdgeMasterSlaveSync
  分类   Category   : DL_Base
  复杂度 Complexity  : cx4
  版本   Version    : 1.0.0
  功能   Purpose    : 主从双通道沿同步判定。主通道越阈上升沿开启 tSyncWindow 等
                      从窗；从沿落在窗内（含与主沿同拍）判通道一致，出单拍有效
                      脉冲；窗内多个从沿只受理第一个；任一信号非有限拍出无效并
                      冻结判定。用于安全回路双通道一致性监视。
  来源   Source     : iec-std-wrapper（T0）
  溯源   Origin     : IEC 61131-3 标准语义的道莅防御性实现；双通道沿一致窗为公开
                      安全仪表语义，clean-room 自研实现，未复制任何闭源代码行。
  平台   Platform   : 纯 IEC 61131-3（TON，无私有库）
  分工声明 Split     : 与 FB_DL_SignalDebounce（单通道消抖）及 FB_DL_Vote2oo3
                      （三选二表决）分工——本件只做双通道沿时序一致性判定，
                      不消抖、不表决、不裁决通道权重。
  作者   Author     : 道莅代码库 · PLC 编程专家（R57）
  ------------------------------------------------------------------
  边界 Boundary     :
                      一 tSyncWindow 钳位 [T#1MS, T#1S]，越界按边界执行并置信息级；
                      二 主从沿同拍判有效（同拍双沿直接出脉冲，不等窗）；
                      三 窗内多从沿只受理第一个（受理即关窗）；
                      四 非有限输入拍：bInvalid 置位、等从窗关闭、不产生脉冲，
                         输出冻结（R191 显式声明），恢复拍不回放历史沿；
                      五 无全局变量、无外部变量声明、无物理地址寻址。
  修订记录 Revision  :
    2026-11-21  v1.0.0  R57 首版（批 1 · 序号 2）
  ==================================================================
*)

TYPE E_DL_EmsPhase :
(
    eIdle      := 0,  // 空闲：等主沿 / idle, waiting for the master edge
    eWaitSlave := 10, // 等从窗：主沿已开窗 / waiting for the slave inside the window
    eFault     := 90  // 无效：输入非有限冻结（信息级驻留，非锁存）/ invalid, a non finite input freezes the grading
);
END_TYPE

FUNCTION_BLOCK FB_DL_EdgeMasterSlaveSync
VAR_INPUT
    fMasterVal  : LREAL := 0.0;  // 主通道信号 [工程单位] / the master channel signal [engineering unit]
    fSlaveVal   : LREAL := 0.0;  // 从通道信号 [工程单位] / the slave channel signal [engineering unit]
    fThresh     : LREAL := 1.0;  // 双通道共用越阈判定阈值 [工程单位] / the shared threshold [engineering unit]
    tSyncWindow : TIME := T#20MS; // 主从沿允许时差窗 [毫秒]，钳位 [1毫秒, 1秒] / the allowed master-slave skew window [millisecond], clamped
    bEnable     : BOOL := TRUE;  // 使能，失能即关窗回空闲 [-] / enable, disabling closes the window
    bReset      : BOOL := FALSE; // 复位上升沿清窗与计数 [-] / reset rising edge clears the window and counters
END_VAR
VAR_OUTPUT
    bSyncValid    : BOOL := FALSE; // 同步有效单拍脉冲 [-] / the sync valid one-scan pulse
    bWaitSlave    : BOOL := FALSE; // 等从窗活动指示 [-] / the window active indicator
    bInvalid      : BOOL := FALSE; // 本拍输入无效（判定冻结）[-] / the inputs are void this scan, the grading frozen
    nMatchCnt     : UDINT := 0;    // 同步有效累计次数 [次] / the accumulated match count [count]
    nLateSlaveCnt : UDINT := 0;    // 窗外迟到从沿累计次数 [次] / the late slave edge count outside the window [count]
    uErrorId      : UDINT := 0;    // 信息级码，0 = 正常 / informational code, zero is ok
    bError        : BOOL := FALSE; // 信息级错误标志（每拍重算，非锁存）/ informational flag, recomputed each scan
END_VAR
VAR
    rtReset : R_TRIG; // 复位沿检测，段 0 无条件刷新 / the reset edge, refreshed unconditionally
    tonWin  : TON;    // 等从窗定时器，段 0 无条件刷新 / the slave window timer, refreshed unconditionally
    _ePhase : E_DL_EmsPhase := E_DL_EmsPhase.eIdle; // 内部相位，CASE 唯一写入目标 / internal phase
    _bInit  : BOOL := FALSE; // 首扫初始化完成标志（R310）/ first scan flag
    _bInOk  : BOOL := FALSE; // 双通道信号均有限 [-] / both signals finite
    _bMNow  : BOOL := FALSE; // 主通道越阈电平（当拍）[-] / the master above-threshold level this scan
    _bSNow  : BOOL := FALSE; // 从通道越阈电平（当拍）[-] / the slave above-threshold level this scan
    _bMPrev : BOOL := FALSE; // 主通道越阈电平（上拍）[-] / the master level previous scan
    _bSPrev : BOOL := FALSE; // 从通道越阈电平（上拍）[-] / the slave level previous scan
    _bMPend : BOOL := FALSE; // 主沿待从标记 [-] / the master edge pending flag
    _tWin   : TIME := T#20MS; // 钳位后的同步窗 [毫秒] / the clamped sync window [millisecond]
END_VAR
VAR CONSTANT
    DL_EMS_WIN_MIN : TIME := T#1MS; // 同步窗下钳位 [毫秒] / the window lower clamp [millisecond]
    DL_EMS_WIN_MAX : TIME := T#1S;  // 同步窗上钳位 [毫秒] / the window upper clamp [millisecond]
END_VAR

// 段 0｜定时器与沿检测无条件周期刷新（禁入分支）/ segment 0, unconditional refresh
rtReset(CLK := bReset); // 复位沿 / the reset edge
tonWin(IN := (_ePhase = E_DL_EmsPhase.eWaitSlave), PT := _tWin); // 等从窗，IN 串等从相闸（无效拍相位已回空闲，天然关窗）/ the window gated by the wait phase, the phase already back to idle on an invalid scan

// 段 1｜首扫初始化（R310）：快照取当拍，禁首拍假边沿 / segment 1, first scan initialisation
IF NOT _bInit THEN // 首扫一拍 / the first scan
    _bInit  := TRUE; // 置首扫标志 / raise the first scan flag
    _bMPrev := FALSE; // 越阈电平从 FALSE 起步（首拍不产沿）/ the level starts FALSE, no edge on the first scan
    _bSPrev := FALSE; // 从通道同理 / the same for the slave
END_IF

// 段 2｜复位沿作用域：清窗 / 清计数（两项逐项声明）/ segment 2, reset edge scope
IF rtReset.Q THEN // 复位沿 / the reset edge
    _bMPend := FALSE; // 作用域一：清主沿待从标记 / scope one, clear the pending flag
    nMatchCnt := 0; // 作用域二：清同步计数 / scope two, clear the match counter
    nLateSlaveCnt := 0; // 作用域二：清迟到计数 / scope two, clear the late counter
END_IF

// 段 3｜输入有限性闸（双判据）与阈值组态闸 / segment 3, the finiteness gate and the threshold gate
_bInOk := (fMasterVal = fMasterVal) AND ((fMasterVal - fMasterVal) = (fMasterVal - fMasterVal)) AND (fSlaveVal = fSlaveVal) AND ((fSlaveVal - fSlaveVal) = (fSlaveVal - fSlaveVal)) AND (fThresh = fThresh) AND ((fThresh - fThresh) = (fThresh - fThresh)); // 双信号与阈值有限性 / finiteness of both signals and the threshold
IF NOT _bInOk THEN // 非有限拍 / a non finite scan
    bInvalid := TRUE; // 置无效标志 / raise the invalid flag
    _bMPend  := FALSE; // 关窗（冻结判定，R191）/ close the window, the grading frozen
    _ePhase  := E_DL_EmsPhase.eIdle; // 回空闲驻留（恢复后重新等主沿）/ back to idle, a fresh wait after recovery
    uErrorId := 16#0001_0002; // 信息级：输入非有限 / informational, a non finite input
    bError   := TRUE; // 置信息级标志 / raise the informational flag
    _bMPrev  := FALSE; // 越阈电平冻结为假（恢复拍不回放历史沿）/ the level frozen false, no historical edge replay
    _bSPrev  := FALSE; // 从通道同理 / the same for the slave
    RETURN; // 早退，脉冲出口保持冻结末值 / early return, the pulse outlet frozen
END_IF

// 段 4｜同步窗钳位（信息级）/ segment 4, the window clamp, informational
IF tSyncWindow < DL_EMS_WIN_MIN THEN // 低于下钳位 / below the lower clamp
    _tWin    := DL_EMS_WIN_MIN; // 钳到下限 / clamp to the floor
    uErrorId := 16#0001_0003; // 信息级：窗过小已钳 / informational, a too small window clamped
    bError   := TRUE; // 置信息级标志 / raise the informational flag
ELSIF tSyncWindow > DL_EMS_WIN_MAX THEN // 高于上钳位 / above the upper clamp
    _tWin    := DL_EMS_WIN_MAX; // 钳到上限 / clamp to the ceiling
    uErrorId := 16#0001_0003; // 信息级：窗过大已钳 / informational, a too large window clamped
    bError   := TRUE; // 置信息级标志 / raise the informational flag
ELSE // 域内 / inside the domain
    _tWin    := tSyncWindow; // 直通 / passthrough
    uErrorId := 16#0000_0000; // 正常码 / the ok code
    bError   := FALSE; // 信息级标志清零 / clear the informational flag
END_IF

// 段 5｜越阈电平与沿提取（R_TRIG 语义手工实现，快照末拍推进）/ segment 5, the above-threshold levels and the edges
_bMNow := fMasterVal > fThresh; // 主通道越阈电平 / the master level
_bSNow := fSlaveVal > fThresh; // 从通道越阈电平 / the slave level

// 段 6｜相位机：ENUM + CASE，含 ELSE 非法相位兜底（R128）/ segment 6, the phase machine
CASE _ePhase OF

E_DL_EmsPhase.eIdle: // 空闲相：等主沿 / the idle phase, waiting for the master edge
    IF _bMNow AND (NOT _bMPrev) THEN // 主沿 / the master edge
        IF _bSNow AND (NOT _bSPrev) THEN // 同拍双沿直接判有效（边界二）/ the same-scan dual edges judged valid
            bSyncValid := TRUE; // 出同步脉冲 / raise the sync pulse
            nMatchCnt := nMatchCnt + 1; // 计数推进 / advance the counter
        ELSE // 无同拍从沿 / no same-scan slave edge
            _bMPend := TRUE; // 开等从窗 / open the window
            _ePhase := E_DL_EmsPhase.eWaitSlave; // 迁等从相 / migrate to the wait phase
        END_IF
    ELSIF _bSNow AND (NOT _bSPrev) THEN // 无主沿的孤立从沿（迟到）/ a lone slave edge, late
        nLateSlaveCnt := nLateSlaveCnt + 1; // 迟到计数 / advance the late counter
    END_IF

E_DL_EmsPhase.eWaitSlave: // 等从相：窗内受理第一个从沿（边界三）/ the wait phase, only the first slave edge accepted
    IF _bSNow AND (NOT _bSPrev) THEN // 从沿到达 / a slave edge arrived
        bSyncValid := TRUE; // 出同步脉冲 / raise the sync pulse
        nMatchCnt := nMatchCnt + 1; // 计数推进 / advance the counter
        _bMPend := FALSE; // 受理即关窗（后续从沿不再受理）/ close on acceptance, later edges not accepted
        _ePhase := E_DL_EmsPhase.eIdle; // 回空闲相 / back to idle
    ELSIF tonWin.Q THEN // 窗满无从沿 / the window expired without a slave edge
        _bMPend := FALSE; // 关窗 / close the window
        _ePhase := E_DL_EmsPhase.eIdle; // 回空闲相 / back to idle
    END_IF

E_DL_EmsPhase.eFault: // 无效驻留相：由段 3 早退覆盖，此处仅兜底 / the invalid dwell phase, covered by the segment three early return
    _ePhase := E_DL_EmsPhase.eIdle; // 兜底回空闲 / fallback to idle

ELSE // 非法相位兜底（R128）/ the illegal phase fallback
    _bMPend := FALSE; // 关窗 / close the window
    _ePhase := E_DL_EmsPhase.eIdle; // 回空闲相 / back to idle
    uErrorId := 16#0001_0005; // 信息级：非法相位 / informational, an illegal phase
    bError   := TRUE; // 置信息级标志 / raise the informational flag
END_CASE

// 段 7｜快照推进与统一出口 / segment 7, the snapshot advance and the unified outlet
_bMPrev := _bMNow; // 主通道快照推进 / advance the master snapshot
_bSPrev := _bSNow; // 从通道快照推进 / advance the slave snapshot
IF NOT _bInOk THEN // 兜底防御（正常路径早退不可达）/ a defensive fallback, unreachable on the normal path
    bSyncValid := FALSE; // 脉冲冻结为假 / the pulse frozen false
END_IF
bWaitSlave := _bMPend; // 等从窗指示 / the window indicator
END_FUNCTION_BLOCK

(* ---- FB_DL_EdgeOrderCheck.st ---- *)
(*==============================================================================
 * 组件名称 (Component)  : FB_DL_EdgeOrderCheck
 * 所属子库 (Sublibrary) : DL_Base
 * 当前版本 (Version)    : 1.0.0
 * 兼容性   (Platform)   : CODESYS 3.5+ / TwinCAT 3 / 汇川 InoProShop / 施耐德 Machine Expert
 *                         仅依赖 Standard.library（TON / R_TRIG / ABS），零厂商私有库
 * 功能描述 (Function)   : 两信号 A→B 时序联锁监视：A 必须先于 B 到达，且 A 领先量
 *                         不少于 tMinGap。逐拍判定四类事件：
 *                         ① 正常顺序：B 上升沿时 A 已在位且领先量 >= tMinGap → bOrderOk TRUE；
 *                         ② 间隔不足：B 上升沿时 A 在位但领先量 < tMinGap → 故障级归因 eGapShort；
 *                         ③ 越序：B 上升沿时 A 不在位（B 无 A 前导）→ 故障级归因 eOrder；
 *                         ④ 逆序：B 先到且仍高，A 随后到来 → nReverseCount 递增并锁存故障 eReverse；
 *                         ⑤ 缺回应：A 单独在位超过 tAloneMax 仍未等到 B → 信息级（不锁故障）。
 * 接口     (Interface)  : 输入 bSigA / bSigB 两信号、tMinGap 最小领先间隔、tAloneMax A 单独
 *                         在位上限、bReset 复位电平；输出 bOrderOk 顺序合规镜像、nReverseCount
 *                         逆序累计计数、eState 相位、eCause 成因、bError、nErrId。
 * 边界     (Boundary)   : ① 组态闸：tMinGap <= T#0S 或 tAloneMax <= tMinGap → 故障锁存；
 *                         ② 计数器饱和于 DL_COUNT_MAX 常量（2147483000，留加 1 裕度，不裸数），
 *                            饱和后不再递增（不回绕，避免台账出现负数）并置信息级留痕；
 *                         ③ R_TRIG 两枚 + TON 两枚在段 0 无条件周期刷新，IN 由当拍电平派生；
 *                         ④ 领先量判据读「前拍快照」_bGapMet：B 上升沿当拍 tonGap.IN 已落假，
 *                            Q 会同拍复位，直接读 Q 会结构性漏判（R45 规则 1 ② 同源教训）；
 *                         ⑤ 故障相迁出唯一路径 = bReset 上升沿；⑥ 零全局耦合（无 GVL / 无物理地址）。
 * 解除式   (Release)    : bReset 上升沿 ∧ 组态合法 ∧ bSigA = FALSE ∧ bSigB = FALSE
 *                         （两信号均已回落，全为当拍量，R240 范式）。自证可满足（终审两式 1）：
 *                         解除式不含任何计时器输出，两信号回落即可达，无恒假因子。
 * 码表     (Codes)      : 16#0001_03EB 故障级：时序联锁故障总码（组态非法 / 间隔不足 / 越序 /
 *                         逆序 / 非法相位），锁存至 bReset 上升沿，归因由 eCause 承载；
 *                         16#0001_04AE 信息级：非故障台账事件（A 缺回应 或 逆序计数饱和）。
 *                         加码反证（R90）：缺回应与计数饱和均不改变 bOrderOk / bError / eCause，
 *                         也无专属状态位可观测，故须立一码留痕；二者共用一码的处置依据是
 *                         「都只要求留痕不要求区分动作」，需要区分时由上层比较
 *                         nReverseCount 是否已达饱和常量反推，无需第二码位。
 *                         码段说明：0001 段故障子带 03xx / 信息子带 04xx，本件取 03EB / 04AE
 *                         （源码实扫该两槽为空，续接同子带已用最大值，未回填碎片孔洞）。
 * 开源溯源 (Origin)     : 道莅自研 clean-room（参考现场联锁惯例与参数域，零代码行复制）
 * 修订历史 (Revision)   : 2026-11-19  v1.0.0  R45 首版（批次 1 · 序号 2）
 *==============================================================================*)

TYPE E_DL_EocState :
(
    eIdle  := 0,     // 双信号均低，等待首个事件 / Idle, both signals low
    eRun   := 10,    // 监视运行（至少一路信号在位） / Running, at least one signal active
    eFault := 90     // 故障锁存相 / Fault latched phase
);
END_TYPE

TYPE E_DL_EocCause :
(
    eNone       := 0,   // 无故障成因 / No cause
    eCfgIllegal := 1,   // 组态非法 / Illegal configuration
    eGapShort   := 2,   // 领先间隔不足 / Lead gap too short
    eOrder      := 3,   // 越序（B 无 A 前导） / Out of order, B without preceding A
    eReverse    := 4    // 逆序（B 先到后 A 到达） / Reverse order, B first then A
);
END_TYPE

FUNCTION_BLOCK FB_DL_EdgeOrderCheck
VAR_INPUT
    bSigA     : BOOL := FALSE;          // 领先信号 A（应先到） [-] / Leading signal A, must arrive first
    bSigB     : BOOL := FALSE;          // 跟随信号 B（应后到） [-] / Following signal B, must arrive later
    tMinGap   : TIME := T#50MS;         // A 领先 B 的最小间隔，域 > T#0S [ms] / Minimum A-to-B lead gap
    tAloneMax : TIME := T#2S;           // A 单独在位上限（缺回应判据），域 > tMinGap [ms] / Max A-alone duration
    bReset    : BOOL := FALSE;          // 复位命令，上升沿清故障 [-] / Reset command, rising edge clears fault
END_VAR
VAR_OUTPUT
    bOrderOk      : BOOL;               // 顺序合规镜像（最近一次 B 沿判定结果） [-] / Order compliance mirror
    nReverseCount : DINT;               // 逆序累计计数（锁存量，复位不清零） [次] / Reverse count, latched, not cleared by reset
    eState        : E_DL_EocState;      // 状态出口，段 6 单点映射 / State outlet
    eCause        : E_DL_EocCause;      // 故障成因出口（R190 归因唯一） / Fault cause outlet
    bError        : BOOL;               // 故障锁存标志 [-] / Fault latch flag
    nErrId        : UDINT;              // 事件码，0 = 无事件 / Event code, 0 = no event
END_VAR
VAR
    _eState       : E_DL_EocState := E_DL_EocState.eIdle;   // 内部相位（CASE 唯一写入目标） / Internal phase
    _eCause       : E_DL_EocCause := E_DL_EocCause.eNone;   // 故障成因锁存（锁存量） / Latched cause
    tonGap        : TON;                // A 领先量计时，段 0 无条件调用 / A lead-gap timer
    tonAlone      : TON;                // A 单独在位计时，段 0 无条件调用 / A-alone duration timer
    rtA           : R_TRIG;             // A 上升沿实例，段 0 无条件调用 / A rising edge
    rtB           : R_TRIG;             // B 上升沿实例，段 0 无条件调用 / B rising edge
    rtReset       : R_TRIG;             // 复位沿实例，段 0 无条件调用 / Reset edge
    _bAlone       : BOOL;               // A 在位且 B 不在位当拍量 [-] / A active while B inactive
    _bGapMet      : BOOL;               // 领先量已满足的前拍快照 [-] / Previous-scan lead-gap satisfied snapshot
    _bCfgBad      : BOOL;               // 组态非法当拍量 [-] / Illegal configuration
    _bFault       : BOOL;               // 故障锁存位（锁存量） / Latched fault bit
    _bOrderOk     : BOOL;               // 顺序合规内部判定（锁存量，供出口映射） / Internal order verdict
    _nReverseCount : DINT;              // 逆序计数内部累计（锁存量，唯一写入点） [次] / Internal reverse counter, single write point [count]
    _uFault       : UDINT;              // 故障码锁存（锁存量） / Latched fault code
    _uInfo        : UDINT;              // 信息码，每拍重算 / Info code, recomputed each scan
END_VAR
VAR CONSTANT
    DL_COUNT_MAX  : DINT := 2147483000; // 逆序计数饱和上限，留安全裕度防加 1 溢出 [次] / Reverse count saturation limit with overflow margin [count]
END_VAR

(* —— 段 0：前拍快照 + 当拍量派生 + 定时器与沿实例无条件周期刷新 —— *)
_bGapMet := tonGap.Q;                                                    // 领先量满足态的前拍快照（B 沿当拍 IN 已落假） / Previous-scan gap-met snapshot
_bAlone  := bSigA AND (NOT bSigB);                                       // A 单独在位当拍量 / A alone this scan
_bCfgBad := (tMinGap <= T#0S) OR (tAloneMax <= tMinGap);                 // 组态非法当拍量 / Illegal configuration
rtA(CLK := bSigA);                                                       // A 上升沿，每拍必调（R228A） / A rising edge, called every scan
rtB(CLK := bSigB);                                                       // B 上升沿，每拍必调 / B rising edge, called every scan
rtReset(CLK := bReset);                                                  // 复位沿，每拍必调 / Reset edge, called every scan
tonGap(IN := _bAlone, PT := tMinGap);                                    // 领先量计时 / Lead-gap timer
tonAlone(IN := _bAlone, PT := tAloneMax);                                // A 单独在位计时 / A-alone timer

(* —— 段 1：单拍量预清零（锁存量与快照量不入清单，R107） —— *)
_uInfo    := 16#0000_0000;         // 信息码每拍重算 / Info recomputed every scan
nErrId    := 16#0000_0000;         // 事件码缺省无事件 / Event code default none
bError    := FALSE;                // 故障标志每拍预清，由故障分支同拍置位（R45 配对） / Flag preset
bOrderOk  := _bOrderOk;            // 顺序镜像由锁存判定派生（名实同源，R191） / Order mirror from latched verdict

(* —— 段 2：复位沿 + 组态域闸 —— *)
IF rtReset.Q THEN                                                        // 当拍复位沿 / current-scan reset edge
    _bFault := FALSE;                                                    // 清故障锁存位（锁存量） / Clear fault latch
    _uFault := 16#0000_0000;                                             // 清故障锁存码（锁存量） / Clear latched code
    _eCause := E_DL_EocCause.eNone;                                      // 清成因（锁存量） / Clear latched cause
    IF _eState = E_DL_EocState.eFault THEN
        _eState := E_DL_EocState.eIdle;                                  // 故障相迁出唯一路径 / Sole exit from fault phase
    END_IF
END_IF
IF _bCfgBad THEN                                                         // 组态域闸 / Configuration gate
    _uFault := 16#0001_03EB;                                             // 故障级：时序联锁故障总码 / Fault-level: order-check fault code
    _bFault := TRUE;                                                     // 锁存置位 / Latch set
    bError  := TRUE;                                                     // 故障标志同拍置位（R45 配对） / Error flag set same scan
    _eCause := E_DL_EocCause.eCfgIllegal;                                // 归因：组态非法 / Cause: illegal configuration
END_IF

(* —— 段 3：顺序判据（B 沿受理 / A 沿逆序判定 / 缺回应信息级） —— *)
IF (NOT _bFault) AND rtB.Q THEN                                          // B 上升沿受理 / B rising edge accepted
    IF bSigA THEN                                                        // A 仍在位：检查领先量 / A is active, check lead gap
        IF _bGapMet THEN
            _bOrderOk := TRUE;                                           // 顺序合规（锁存量） / Order OK, latched verdict
        ELSE
            _uFault := 16#0001_03EB;
            _bFault := TRUE;
            bError  := TRUE;
            _eCause := E_DL_EocCause.eGapShort;                          // 归因：领先间隔不足 / Cause: lead gap too short
            _bOrderOk := FALSE;                                          // 锁存量置违规 / Latched verdict violation
        END_IF
    ELSE
        _uFault := 16#0001_03EB;
        _bFault := TRUE;
        bError  := TRUE;
        _eCause := E_DL_EocCause.eOrder;                                 // 归因：越序（B 无 A 前导） / Cause: out of order
        _bOrderOk := FALSE;                                              // 锁存量置违规 / Latched verdict violation
    END_IF
END_IF
IF (NOT _bFault) AND rtA.Q AND bSigB THEN                                // A 在 B 仍高时到来 = 逆序 / A arrives while B still high
    IF _nReverseCount < DL_COUNT_MAX THEN
        _nReverseCount := _nReverseCount + 1;                            // 逆序计数递增（单点写入） / Reverse count increment, single write point
    ELSE
        _uInfo := 16#0001_04AE;                                          // 信息级：计数饱和留痕，不回绕 / Info: saturation recorded, no wrap
    END_IF
    _uFault := 16#0001_03EB;
    _bFault := TRUE;
    bError  := TRUE;
    _eCause := E_DL_EocCause.eReverse;                                   // 归因：逆序 / Cause: reverse order
    _bOrderOk := FALSE;                                                  // 锁存量置违规 / Latched verdict violation
END_IF
IF (NOT _bFault) AND tonAlone.Q THEN                                     // A 单独在位超上限 → 缺回应（信息级，不锁故障） / A alone too long, info level
    _uInfo := 16#0001_04AE;
END_IF

(* —— 段 4：故障解除式（R240 全当拍量） —— *)
IF rtReset.Q AND (NOT _bCfgBad) AND (NOT bSigA) AND (NOT bSigB) THEN
    _bFault := FALSE;                                                    // 清故障锁存位（锁存量） / Clear fault latch
    _uFault := 16#0000_0000;                                             // 清故障锁存码（锁存量） / Clear latched code
    _eCause := E_DL_EocCause.eNone;                                      // 清成因（锁存量） / Clear latched cause
END_IF

(* —— 段 4A：故障锁存相位迁移闸 —— *)
IF _bFault AND (_eState <> E_DL_EocState.eFault) THEN
    _eState := E_DL_EocState.eFault;                                     // 锁存即入故障相 / Latch enters fault phase
END_IF

(* —— 段 5：相位机（ENUM 全成员显式标签 + ELSE 兜底，R128） —— *)
CASE _eState OF

E_DL_EocState.eIdle:
    IF bSigA OR bSigB THEN                                               // 出口 1：任一信号动作 / Any signal active
        _eState := E_DL_EocState.eRun;
    ELSIF _bFault THEN                                                   // 出口 2：故障锁存 / Fault latched
        _eState := E_DL_EocState.eFault;
    END_IF

E_DL_EocState.eRun:
    IF (NOT bSigA) AND (NOT bSigB) THEN                                  // 出口 1：两信号均回落 / Both signals released
        _eState := E_DL_EocState.eIdle;
    ELSIF _bFault THEN                                                   // 出口 2：故障锁存 / Fault latched
        _eState := E_DL_EocState.eFault;
    END_IF

E_DL_EocState.eFault:
    ;                                                                     // 故障相：仅段 4 复位沿可迁出 / Only the reset edge leaves this phase

ELSE
    _uFault := 16#0001_03EB;                                             // 故障级：非法相位兜底（归并总码） / Illegal-phase fallback
    _bFault := TRUE;
    bError  := TRUE;
    _eCause := E_DL_EocCause.eCfgIllegal;                                // 归因：相位非法归并组态 / Cause: phase illegal
    _eState := E_DL_EocState.eFault;

END_CASE

(* —— 段 6：出口单点映射（名实同源；锁存码回放） —— *)
nReverseCount := _nReverseCount;                                         // 逆序计数出口（锁存量回放） / Reverse count outlet
IF _bFault THEN
    bOrderOk := FALSE;                                                   // 故障相强制违规镜像 / Fault forces violation mirror
    nErrId   := _uFault;                                                 // 故障锁存码回放 / Replay latched fault code
ELSE
    nErrId   := _uInfo;                                                  // 信息码 / Info code
END_IF
bError := _bFault;                                                       // 故障标志与锁存同源（名实双出口，R191） / Flag from latch
eState := _eState;                                                       // 状态出口 / State outlet
eCause := _eCause;                                                       // 成因出口 / Cause outlet

END_FUNCTION_BLOCK

(* ---- FB_DL_EncoderQuadCount.st ---- *)
(*
  ==================================================================
  组件名 Component  : FB_DL_EncoderQuadCount
  分类   Category   : DL_Base
  复杂度 Complexity  : cx5
  版本   Version    : 1.0.1
  功能   Purpose    : 正交 A/B 两相四倍频加减计数。按格雷序四态状态机解码相位
                      跳变方向；A/B 同拍跳变（非法 00↔11 或 01↔10）按状态保持
                      并按 2 步口径累计丢步；计数饱和 ±DL_ENC_QUAD_MAX 口径不回
                      绕；方向出口与计数出口分离。
  来源   Source     : iec-std-wrapper（T0）
  溯源   Origin     : IEC 61131-3 标准语义的道莅防御性实现；正交解码格雷序四态
                      状态机为公开编码器语义，clean-room 自研实现，未复制任何
                      厂商私有库源码。
  平台   Platform   : 纯 IEC 61131-3（无私有库、无定时器实例、无 MOD 于计数路径）
  分工声明 Split     : 与 FB_DL_HistogramAccum / FB_DL_EventRateCalc 分工——本件
                      只做正交相位解码与四倍频计数，不做速率换算与统计分箱。
  作者   Author     : 道莅代码库 · PLC 编程专家（R57）
  ------------------------------------------------------------------
  边界 Boundary     :
                      一 首扫经 _bFirst 豁免一拍步进判定（v1.0.1）：首拍只锁存
                         格雷态，不产生任何计数与方向（消除上电停在非 00 态时
                         用陈旧 _eGrayPv 判转移的首拍假步进）；
                      二 非法跳变（对角跳 00↔11 / 01↔10）状态保持、计数不动、
                         丢步按 2 步口径累计（v1.0.1 A 案：一个对角跳变实际
                         丢失 2 个四分之一周期步，计数单位 [步]）；
                      三 计数饱和 ±DL_ENC_QUAD_MAX，饱和侧锁存指示，不回绕；
                      四 方向出口只随最近一次有效步进更新，非法跳变不改方向；
                      五 无全局变量、无外部变量声明、无物理地址寻址。
  修订记录 Revision  :
    2026-11-21  v1.0.0  R57 首版（批 1 · 序号 3）
    2026-11-21  v1.0.1  R58 返修两项：①段 1 的 _bInit 预置 _eGrayNow 为死代码
                        （当拍即被段 3 重锁存覆盖），改置 _bFirst 豁免首拍步进
                        判定；②丢步判式口径二选一：全库检索无手册引用，选 A
                        案代码改——对角非法跳变按丢失 2 步累计（四分支 + 兜底
                        分支同口径），计数单位 [步]，头注释边界二同步改写。
  ==================================================================
*)

TYPE E_DL_EncGray :
(
    eQ0 := 0, // 格雷态 0：A=0 / B=0（AB 编码 00）/ gray state zero, A low and B low
    eQ1 := 1, // 格雷态 1：A=0 / B=1（AB 编码 01）/ gray state one, A low and B high
    eQ3 := 3, // 格雷态 3：A=1 / B=1（AB 编码 11）/ gray state three, A high and B high
    eQ2 := 2  // 格雷态 2：A=1 / B=0（AB 编码 10）/ gray state two, A high and B low
);
END_TYPE

FUNCTION_BLOCK FB_DL_EncoderQuadCount
VAR_INPUT
    bPhaseA  : BOOL := FALSE;       // 正交 A 相输入 [-] / the quadrature phase A input
    bPhaseB  : BOOL := FALSE;       // 正交 B 相输入 [-] / the quadrature phase B input
    bEnable  : BOOL := TRUE;        // 使能，失能冻结计数 [-] / enable, disabling freezes the count
    bReset   : BOOL := FALSE;       // 复位上升沿清计数与丢步 [-] / reset rising edge clears the count and missed steps
END_VAR
VAR_OUTPUT
    nQuadCount : DINT := 0;   // 四倍频计数出口（饱和 ±上限，不回绕）[步] / the quadrature count outlet, saturated, no wrap [step]
    bDirPos    : BOOL := FALSE; // 方向出口，TRUE = 最近有效步进为正向 [-] / the direction outlet, true for the latest valid forward step
    bSatHi     : BOOL := FALSE; // 正向饱和锁存指示 [-] / the forward saturation latch indicator
    bSatLo     : BOOL := FALSE; // 反向饱和锁存指示 [-] / the reverse saturation latch indicator
    nMissCnt   : UDINT := 0;    // 非法跳变丢步累计（对角跳变按 2 步计，v1.0.1 A 案）[步] / the illegal transition missed count in steps, a diagonal counts two
    bError     : BOOL := FALSE; // 故障标志（保留位，本件无锁存故障）[-] / the fault flag, reserved, no latched fault
END_VAR
VAR
    rtReset   : R_TRIG; // 复位沿检测，段 0 无条件刷新 / the reset edge, refreshed unconditionally
    _eGrayPv  : E_DL_EncGray := E_DL_EncGray.eQ0; // 上拍格雷态 / the previous gray state
    _eGrayNow : E_DL_EncGray := E_DL_EncGray.eQ0; // 当拍格雷态 / the current gray state
    _bInit    : BOOL := FALSE; // 首扫初始化完成标志（R310）/ first scan flag
    _bFirst   : BOOL := FALSE; // 首拍跳过步进判定标记（v1.0.1 豁免一拍）/ the first scan skip flag, exempts one scan
    _nStep    : DINT := 0;     // 本拍步进量（+1、-1、0 三值）[步] / the step amount this scan [step]
    _nMissAdd : DINT := 0;     // 本拍丢步累加量，对角跳变按 2 [步] / the miss addition this scan, a diagonal counts two [step]
END_VAR
VAR CONSTANT
    DL_ENC_QUAD_MAX : DINT := 2147483600; // 四倍频计数饱和上限 [步]，留 47 步余量防 ±1 回绕 / the saturation bound [step], a margin against a plus or minus one wrap
    DL_ENC_MISS_MAX : UDINT := 4294967293; // 丢步计数钳定界 [步]，留 2 步余量防累加回绕 / the missed count clamp [step], a two step margin against a wrap
END_VAR

// 段 0｜沿检测无条件周期刷新（禁入分支）/ segment 0, unconditional refresh
rtReset(CLK := bReset); // 复位沿 / the reset edge

// 段 1｜首扫初始化（R310）：置 _bFirst 豁免一拍，零计数零方向（v1.0.1）/ segment 1, the first scan raises the exemption flag
IF NOT _bInit THEN // 首扫一拍 / the first scan
    _bInit  := TRUE; // 置首扫标志 / raise the first scan flag
    _bFirst := TRUE; // 首拍豁免步进判定（上电停在非 00 态不用陈旧 _eGrayPv 判转移）/ exempt the first scan from the step verdict
END_IF

// 段 2｜复位沿作用域：清计数 / 清方向 / 清饱和与丢步（四项逐项声明）/ segment 2, reset edge scope
IF rtReset.Q THEN // 复位沿 / the reset edge
    nQuadCount := 0; // 作用域一：清计数 / scope one, clear the count
    bDirPos := FALSE; // 作用域二：清方向 / scope two, clear the direction
    bSatHi := FALSE; // 作用域三：清正向饱和 / scope three, clear the forward saturation
    bSatLo := FALSE; // 作用域三：清反向饱和 / scope three, clear the reverse saturation
    nMissCnt := 0; // 作用域四：清丢步计数 / scope four, clear the missed counter
END_IF

// 段 3｜当拍格雷态解码（A 低位 B 高位，纯布尔组合，无 MOD 无移位）/ segment 3, the gray decode, pure boolean composition
_eGrayNow := E_DL_EncGray.eQ0; // 默认态 00 / the default state
IF bPhaseA AND (NOT bPhaseB) THEN _eGrayNow := E_DL_EncGray.eQ2; END_IF // 编码 10 / the encoding ten
IF (NOT bPhaseA) AND bPhaseB THEN _eGrayNow := E_DL_EncGray.eQ1; END_IF // 编码 01 / the encoding one
IF bPhaseA AND bPhaseB THEN _eGrayNow := E_DL_EncGray.eQ3; END_IF // 编码 11 / the encoding eleven

// 段 4｜步进与丢步判定：格雷序状态机 CASE，非法跳变保持丢步（边界二）/ segment 4, the step and miss verdict
_nStep    := 0; // 步进量预置零 / preset the step to zero
_nMissAdd := 0; // 丢步累加量预置零 / preset the miss addition to zero
IF bEnable AND (NOT _bFirst) AND (_eGrayNow <> _eGrayPv) THEN // 使能且非首拍且格雷态变化（v1.0.1 豁免闸）/ enabled, not the first scan, and the gray state changed
    CASE _eGrayPv OF // 以上拍态为基准查转移表 / the transition table keyed by the previous state

    E_DL_EncGray.eQ0: // 上拍 00 / the previous state zero
        IF _eGrayNow = E_DL_EncGray.eQ1 THEN // 00→01 正向四分之一周期 / a forward quarter cycle
            _nStep := 1; // 正向步进 / a forward step
        ELSIF _eGrayNow = E_DL_EncGray.eQ2 THEN // 00→10 反向四分之一周期 / a reverse quarter cycle
            _nStep := -1; // 反向步进 / a reverse step
        ELSE // 00→11 对角非法跳变 / the diagonal illegal transition
            _nMissAdd := 2; // 对角跳变按丢失 2 步计（v1.0.1 A 案）/ a diagonal transition counts as two lost steps
        END_IF

    E_DL_EncGray.eQ1: // 上拍 01 / the previous state one
        IF _eGrayNow = E_DL_EncGray.eQ3 THEN // 01→11 正向 / a forward transition
            _nStep := 1; // 正向步进 / a forward step
        ELSIF _eGrayNow = E_DL_EncGray.eQ0 THEN // 01→00 反向 / a reverse transition
            _nStep := -1; // 反向步进 / a reverse step
        ELSE // 01→10 对角非法 / the diagonal illegal transition
            _nMissAdd := 2; // 对角跳变按丢失 2 步计（v1.0.1 A 案）/ a diagonal transition counts as two lost steps
        END_IF

    E_DL_EncGray.eQ3: // 上拍 11 / the previous state three
        IF _eGrayNow = E_DL_EncGray.eQ2 THEN // 11→10 正向 / a forward transition
            _nStep := 1; // 正向步进 / a forward step
        ELSIF _eGrayNow = E_DL_EncGray.eQ1 THEN // 11→01 反向 / a reverse transition
            _nStep := -1; // 反向步进 / a reverse step
        ELSE // 11→00 对角非法 / the diagonal illegal transition
            _nMissAdd := 2; // 对角跳变按丢失 2 步计（v1.0.1 A 案）/ a diagonal transition counts as two lost steps
        END_IF

    E_DL_EncGray.eQ2: // 上拍 10 / the previous state two
        IF _eGrayNow = E_DL_EncGray.eQ0 THEN // 10→00 正向 / a forward transition
            _nStep := 1; // 正向步进 / a forward step
        ELSIF _eGrayNow = E_DL_EncGray.eQ3 THEN // 10→11 反向 / a reverse transition
            _nStep := -1; // 反向步进 / a reverse step
        ELSE // 10→01 对角非法 / the diagonal illegal transition
            _nMissAdd := 2; // 对角跳变按丢失 2 步计（v1.0.1 A 案）/ a diagonal transition counts as two lost steps
        END_IF

    ELSE // 非法格雷态兜底（R128，实际不可达：_eGrayPv 只取自段 3 四态解码）/ the illegal gray fallback, unreachable since the snapshot only takes the four decoded states
        _nMissAdd := 2; // 兜底与对角跳变同口径按 2 步计（v1.0.1）/ the fallback aligns with the diagonal two step convention
    END_CASE
END_IF
_bFirst := FALSE; // 首拍标记仅豁免一拍（v1.0.1，段 4 之后段 5 之前清除）/ the first scan flag exempts only one scan, cleared after segment four

// 段 5｜饱和计数写入点唯一（净额单点施加，R47）/ segment 5, the single count write point with saturation
IF _nStep > 0 THEN // 正向步进 / a forward step
    IF nQuadCount >= DL_ENC_QUAD_MAX THEN // 已在正向饱和界 / already at the forward bound
        bSatHi := TRUE; // 锁存饱和指示 / latch the saturation indicator
    ELSE // 未饱和 / not saturated
        nQuadCount := nQuadCount + 1; // 计数 +1 / count up
        bDirPos := TRUE; // 方向出口置正 / the direction outlet positive
    END_IF
ELSIF _nStep < 0 THEN // 反向步进 / a reverse step
    IF nQuadCount <= -DL_ENC_QUAD_MAX THEN // 已在反向饱和界 / already at the reverse bound
        bSatLo := TRUE; // 锁存饱和指示 / latch the saturation indicator
    ELSE // 未饱和 / not saturated
        nQuadCount := nQuadCount - 1; // 计数 -1 / count down
        bDirPos := FALSE; // 方向出口置负 / the direction outlet negative
    END_IF
END_IF
IF _nMissAdd > 0 THEN // 非法跳变丢步（状态保持、计数不动、方向不改，边界二四）/ an illegal transition, the state held, the count untouched, the direction unchanged
    nMissCnt := nMissCnt + DINT_TO_UDINT(_nMissAdd); // 丢步累计按步口径推进（v1.0.1 A 案）/ advance the missed count in steps
    IF nMissCnt > DL_ENC_MISS_MAX THEN // UDINT 上界防回绕（钳定界留 2 步累加余量）/ the wrap guard clamped with a two step margin
        nMissCnt := DL_ENC_MISS_MAX; // 钳在安全界 / clamp below the ceiling
    END_IF
END_IF

// 段 6｜格雷态快照推进（无条件，失能拍也推进防恢复假跳变）/ segment 6, the gray snapshot advances unconditionally
_eGrayPv := _eGrayNow; // 快照推进 / advance the snapshot
END_FUNCTION_BLOCK

(* ---- FB_DL_EStopDualChannel.st ---- *)
(*
  ==================================================================
  组件名 Component  : FB_DL_EStopDualChannel
  分类   Category   : DL_Base
  复杂度 Complexity  : cx4
  版本   Version    : 1.0.0
  功能   Purpose    : 双通道急停监视。两路常闭信号（TRUE = 触点闭合 = 安全侧）做
                      一致性监视：两路均闭合出安全态；仅一路闭合进入差异窗
                      （tDiscMax），超窗判单通道失效并锁存坏通道位；两路均断开
                      判「已拍下」（信息级，安全侧输出为假）；复位上升沿必须在
                      两通道均恢复后到达才可清锁存，未恢复即按复位判 eStuckReset。
  来源   Source     : t2-1-lgf-converter（安全逻辑组织）
  溯源   Origin     : IEC 61131-3 标准语义的道莅防御性实现；双回路不一致监视组织
                      借鉴 IEC 60204-1 公开条款语义，clean-room 自研，未复制任何
                      闭源代码行。
  平台   Platform   : 纯 IEC 61131-3（TON / R_TRIG，无私有库）
  作者   Author     : 道莅代码库 · PLC 编程专家（R56）
  ------------------------------------------------------------------
  边界 Boundary     :
                      一 本件只做双回路监视与安全侧出口，不驱动任何执行器（属主边界）；
                      二 bSafeState 只在两通道均确认安全（均闭合）且无故障锁存时为真，
                         任何不确定一律走 FALSE（安全侧优先，失效即断开语义）；
                      三 eBothOpen 为信息级成因（正常拍下状态），不置 bError；
                         其余成因均为故障级，与 bError 配对（R45）；
                      四 故障锁存解除路径 = bReset 上升沿且两通道均闭合（唯一路径，
                         头注释声明，R188）；未恢复即复位判 eStuckReset 并锁存；
                      五 差异自愈：差异窗内两通道恢复一致即回运行相，不锁存（瞬时抖动
                         不判失效，tDiscMax 内自愈为设计意图）；
                      六 无全局变量、无外部变量声明、无物理地址寻址。
  输出契约 Output contract:
                      bChannel1Bad / bChannel2Bad 为锁存位，仅在 eDiscTimeout 判定时
                      置位（坏通道 = 处于断开位的那一路），复位沿恢复后清零；
                      eFault 为锁存回放（不在故障相按当下输入重推断，R152）；
                      ePhaseBad 为非法相位兜底专用成员（R128）。
  修订记录 Revision  :
    2026-11-20  v1.0.0  R56 首版（批 1 · 序号 5）
  ==================================================================
*)

TYPE E_DL_EsdPhase :
(
    eIdle    := 0,  // 未使能：监视停摆，安全侧输出为假 / disabled, the watch is idle and the safe outlet is false
    eRun     := 10, // 运行：两通道一致（均闭合或均断开）/ running, the channels agree
    eDiscord := 20, // 差异：仅一路闭合，差异窗计时中 / discrepancy, one channel closed and the window is timing
    eFault   := 90  // 故障：成因锁存，安全侧输出为假 / fault, the cause is latched and the safe outlet is false
);
END_TYPE

TYPE E_DL_EsdFault :
(
    eNone            := 0, // 无成因 / no cause
    eChannelMismatch := 1, // 通道不一致（差异窗内，信息级）/ the channels disagree inside the window, informational
    eDiscTimeout     := 2, // 差异超窗判单通道失效（故障级，与 bError 配对）/ the discrepancy outlasted the window, a single channel failed, fault grade paired with bError
    eBothOpen        := 3, // 两路均断开 = 急停已拍下（信息级，安全侧为假）/ both channels open, the stop is pressed, informational
    eStuckReset      := 4, // 复位到达但通道未恢复（故障级，与 bError 配对）/ a reset arrived without both channels restored, fault grade paired with bError
    ePhaseBad        := 5  // 非法相位兜底（故障级，与 bError 配对）/ illegal phase fallback, fault grade paired with bError
);
END_TYPE

FUNCTION_BLOCK FB_DL_EStopDualChannel
VAR_INPUT
    bEnable  : BOOL := TRUE;      // 使能，失能时安全侧输出为假 [-] / enable, the safe outlet is false when disabled
    bReset   : BOOL := FALSE;     // 复位，上升沿在两通道均闭合时清锁存 [-] / reset, the rising edge clears the latch only with both channels closed
    bCh1Ok   : BOOL := TRUE;      // 通道 1 常闭反馈，TRUE = 闭合 = 安全 [-] / channel one normally closed feedback, true is closed and safe
    bCh2Ok   : BOOL := TRUE;      // 通道 2 常闭反馈，TRUE = 闭合 = 安全 [-] / channel two normally closed feedback, true is closed and safe
    tDiscMax : TIME := T#500MS;   // 差异窗（单通道失效判定时长）[毫秒]，域 大于零 / discrepancy window [millisecond], domain above zero
END_VAR
VAR_OUTPUT
    bSafeState    : BOOL := FALSE; // 安全侧输出：仅在两通道均闭合且无故障锁存时为真 [-] / the safe side outlet, true only with both channels closed and no fault latch
    bChannel1Bad  : BOOL := FALSE; // 通道 1 失效锁存位 [-] / channel one failed latch bit
    bChannel2Bad  : BOOL := FALSE; // 通道 2 失效锁存位 [-] / channel two failed latch bit
    ePhase        : E_DL_EsdPhase := E_DL_EsdPhase.eIdle; // 相位出口 [枚举] / phase outlet [enum]
    eFault        : E_DL_EsdFault := E_DL_EsdFault.eNone; // 成因出口，锁存回放 [枚举] / cause outlet replayed from the latch [enum]
    bError        : BOOL := FALSE; // 故障锁存标志 [-] / fault latch flag
END_VAR
VAR
    rtReset  : R_TRIG; // 复位沿检测，段 0 无条件刷新 / reset edge detector, refreshed unconditionally in segment zero
    tonDisc  : TON;    // 差异窗计时，段 0 无条件刷新 / discrepancy window timer, refreshed unconditionally in segment zero
    _ePhase  : E_DL_EsdPhase := E_DL_EsdPhase.eIdle; // 内部相位，CASE 唯一写入目标 / internal phase, the only CASE write target
    _eCause  : E_DL_EsdFault := E_DL_EsdFault.eNone; // 信息级成因，每拍重算 / informational cause, recomputed every scan
    _eFaulC  : E_DL_EsdFault := E_DL_EsdFault.eNone; // 故障级成因，锁存至复位沿 / fault cause, latched until the reset edge
    _bFault  : BOOL := FALSE; // 故障锁存位 [-] / fault latch bit
    _bInit   : BOOL := FALSE; // 首扫初始化完成标志（R310）/ first scan initialisation flag
    _bDisc   : BOOL := FALSE; // 本拍通道不一致 [-] / the channels disagree this scan
    _bBothOk : BOOL := FALSE; // 本拍两通道均闭合 [-] / both channels are closed this scan
    _bNoneOk : BOOL := FALSE; // 本拍两通道均断开 [-] / both channels are open this scan
END_VAR

// 段 0｜定时器与沿检测无条件周期刷新（禁入分支），IN 只串相位闸与故障闸 / segment 0, unconditional refresh with the phase and fault gates on IN only
rtReset(CLK := bReset); // 复位沿无条件刷新 / unconditional refresh of the reset edge
tonDisc(IN := (_ePhase = E_DL_EsdPhase.eDiscord) AND (NOT _bFault), PT := tDiscMax); // 差异窗，IN 串差异相闸与故障闸 / the discrepancy window with the phase and fault gates on IN

// 段 1｜首扫初始化（R310）/ segment 1, first scan initialisation
IF NOT _bInit THEN // 首扫一拍 / the very first scan
    _bInit := TRUE; // 置首扫完成标志 / raise the first scan flag
    _ePhase := E_DL_EsdPhase.eRun; // 相位从运行起步（使能默认真）/ the phase starts in run
    _eCause := E_DL_EsdFault.eNone; // 信息级成因清零 / clear the informational cause
    _eFaulC := E_DL_EsdFault.eNone; // 故障级成因清零 / clear the fault cause
    _bFault := FALSE; // 故障锁存清零 / clear the fault latch
END_IF

// 段 2｜本拍一致性判定（组合量，无锁存）/ segment 2, the per scan consistency verdict
_bBothOk := bCh1Ok AND bCh2Ok; // 两路均闭合 / both channels are closed
_bNoneOk := (NOT bCh1Ok) AND (NOT bCh2Ok); // 两路均断开 / both channels are open
_bDisc := (bCh1Ok <> bCh2Ok); // 两路不一致（XOR 语义）/ the channels disagree

// 段 3｜复位沿作用域：仅在两通道均恢复时清锁存，未恢复判卡死复位 / segment 3, reset edge scope, the latch clears only with both channels restored
IF rtReset.Q THEN // 复位沿 / the reset edge
    IF _bBothOk THEN // 两通道均恢复 / both channels are restored
        _bFault := FALSE; // 作用域一：清故障锁存 / scope one, clear the fault latch
        _eFaulC := E_DL_EsdFault.eNone; // 作用域一：清故障级成因 / scope one, clear the fault cause
        bChannel1Bad := FALSE; // 作用域一：清通道 1 失效位 / scope one, clear the channel one failed bit
        bChannel2Bad := FALSE; // 作用域一：清通道 2 失效位 / scope one, clear the channel two failed bit
        _ePhase := E_DL_EsdPhase.eRun; // 作用域二：迁回运行相 / scope two, migrate back to run
    ELSE // 未恢复即复位 / a reset without restoration
        _bFault := TRUE; // 置故障锁存 / raise the fault latch
        _eFaulC := E_DL_EsdFault.eStuckReset; // 故障级成因（R45 配对 bError）/ the fault cause paired with bError
        _ePhase := E_DL_EsdPhase.eFault; // 迁故障相 / migrate to the fault phase
    END_IF
END_IF

// 段 4｜相位机：ENUM + CASE，含 ELSE 非法相位兜底（R128）/ segment 4, the phase machine with an ELSE fallback
CASE _ePhase OF
E_DL_EsdPhase.eIdle: // 未使能相：安全侧输出为假 / the disabled phase, the safe outlet is false
    IF bEnable THEN // 使能恢复 / enabled again
        _ePhase := E_DL_EsdPhase.eRun; // 迁运行相 / migrate to run
    END_IF

E_DL_EsdPhase.eRun: // 运行相：两通道一致 / the run phase, the channels agree
    IF NOT bEnable THEN // 失能 / disabled
        _ePhase := E_DL_EsdPhase.eIdle; // 迁未使能相 / migrate to idle
    ELSIF _bDisc THEN // 通道不一致 / the channels disagree
        _eCause := E_DL_EsdFault.eChannelMismatch; // 信息级成因：差异窗内 / the informational cause inside the window
        _ePhase := E_DL_EsdPhase.eDiscord; // 迁差异相 / migrate to the discrepancy phase
    ELSIF _bNoneOk THEN // 两路均断开 = 已拍下 / both open, the stop is pressed
        _eCause := E_DL_EsdFault.eBothOpen; // 信息级成因，不置故障（设计语义）/ the informational cause, no fault by design
    ELSE // 两路均闭合，无成因 / both closed, no cause
        _eCause := E_DL_EsdFault.eNone; // 成因清零 / clear the cause
    END_IF

E_DL_EsdPhase.eDiscord: // 差异相：差异窗计时 / the discrepancy phase, the window is timing
    IF NOT bEnable THEN // 失能 / disabled
        _ePhase := E_DL_EsdPhase.eIdle; // 迁未使能相 / migrate to idle
    ELSIF _bBothOk THEN // 差异自愈：窗内恢复一致（R152 自愈路径）/ the transient self heals inside the window
        _eCause := E_DL_EsdFault.eNone; // 成因清零 / clear the cause
        _ePhase := E_DL_EsdPhase.eRun; // 迁回运行相 / migrate back to run
    ELSIF _bNoneOk THEN // 两路均断开，回到一致（已拍下）/ both open, consistent again
        _eCause := E_DL_EsdFault.eBothOpen; // 信息级成因 / the informational cause
        _ePhase := E_DL_EsdPhase.eRun; // 迁回运行相 / migrate back to run
    ELSIF tonDisc.Q THEN // 差异超窗：判单通道失效 / the window expired, a single channel failed
        bChannel1Bad := NOT bCh1Ok; // 坏通道 1 = 处于断开位的一路 / channel one is bad when it sits open
        bChannel2Bad := NOT bCh2Ok; // 坏通道 2 同口径 / channel two the same way
        _bFault := TRUE; // 置故障锁存 / raise the fault latch
        _eFaulC := E_DL_EsdFault.eDiscTimeout; // 故障级成因（R45 配对 bError）/ the fault cause paired with bError
        _ePhase := E_DL_EsdPhase.eFault; // 迁故障相 / migrate to the fault phase
    ELSE // 差异仍在窗内 / the discrepancy persists inside the window
        _eCause := E_DL_EsdFault.eChannelMismatch; // 信息级成因每拍重算 / the informational cause is recomputed every scan
    END_IF

E_DL_EsdPhase.eFault: // 故障相：成因锁存回放，安全侧输出为假 / the fault phase, the cause is latched and the safe outlet is false
    IF NOT bEnable THEN // 失能 / disabled
        _ePhase := E_DL_EsdPhase.eIdle; // 迁未使能相 / migrate to idle
    END_IF

ELSE // 非法相位兜底（R128）/ the illegal phase fallback
    _bFault := TRUE; // 置故障锁存 / raise the fault latch
    _eFaulC := E_DL_EsdFault.ePhaseBad; // 故障级成因（R45 配对 bError）/ the fault cause paired with bError
    _ePhase := E_DL_EsdPhase.eFault; // 迁故障相 / migrate to the fault phase
END_CASE

// 段 5｜统一出口：安全侧出口与成因锁存回放 / segment 5, the unified outlet with the safe side and the latched cause
IF _bFault THEN // 故障锁存优先 / the fault latch takes priority
    eFault := _eFaulC; // 故障级成因锁存回放（不按当下输入重推断，R152）/ the fault cause replayed from the latch
ELSE
    eFault := _eCause; // 信息级成因直映 / the informational cause is mapped directly
END_IF
bSafeState := bCh1Ok AND bCh2Ok AND (NOT _bFault) AND bEnable; // 安全侧出口：双确认 + 无锁存 + 使能（任何不确定走假）/ the safe outlet, double confirmation without a latch, any doubt is false
ePhase := _ePhase; // 相位出口单点映射 / single point phase outlet mapping
bError := _bFault; // 故障标志与锁存位同源 / the fault flag shares the latch source
END_FUNCTION_BLOCK
